// ---- 20_Module/Mqtt/Config/ST_ScheduleWeekly_V1.TcDUT
{attribute 'pack_mode' := '1'}
TYPE ST_ScheduleWeekly_V1 :
STRUCT
 Name : STRING(20);
 Priority : UDINT;
 StartDate : UDINT;
 EndDate : UDINT;
 Works : ARRAY[0..69] OF ST_ScheduleWork_V1;
END_STRUCT
END_TYPE

// ---- 20_Module/Mqtt/ST_IfUpsConfigRx.TcDUT
// MQTT로 받은 UPS 설정을 프로그램에 넘기는 묶음.
// 현재 수신만 하고 장비에는 적용하지 않는다.
{attribute 'pack_mode' := '1'}
TYPE ST_IfUpsConfigRx :
STRUCT
 nRxCount : UDINT; // 수신 누계
 astConfig : ARRAY[0..GVL_PARAM.UPS_COUNT-1] OF ST_UpsConfig_Rx; // UPS별 설정
END_STRUCT
END_TYPE

// ---- 20_Module/Ups/E_UpsChargeAction.TcDUT
// 충방전 시퀀스가 요청하는 동작. ST_UpsChargeRequest.eAction에 담긴다.
{attribute 'qualified_only'}
{attribute 'strict'}
TYPE E_UpsChargeAction : (
 NoRequest := 0, // 요청 없음
 BbcOn := 1, // BBC 기동
 BbcReady := 2, // BBC 대기 (현재 맵에 명령 없음, 확인 필요)
 BmsPreparePeriodic := 3, // BMS 주기적 방전 준비
 BmsPreparePulse := 4, // BMS 펄스 방전 준비
 PeriodicStart := 5, // UPS 주기적 방전 시작
 PulseStart := 6, // UPS 펄스 방전 시작
 DischargeCancel := 7, // UPS 방전 취소
 BmsDischargeCancel := 8, // BMS 방전 취소
 FloatCharge := 9, // 부동충전 복귀
 ChargeVoltage := 10 // 충전 전압 적용 (온도보상, fValue 사용)
) INT;
END_TYPE

// ---- 20_Module/Ups/E_UpsChargeMode.TcDUT
// 충방전 시퀀스의 운전 종류. 주 운전이라 한 번에 하나만 실행한다.
{attribute 'qualified_only'}
{attribute 'strict'}
TYPE E_UpsChargeMode : (
 Off := 0, // 운전 없음
 Trickle := 1, // 간헐충전
 Periodic := 2, // 주기적 방전
 Pulse := 3 // 펄스 방전
) INT;
END_TYPE

// ---- 20_Module/Ups/E_UpsChargeStep.TcDUT
// FB_UpsChargeSequence의 진행 단계.
{attribute 'qualified_only'}
{attribute 'strict'}
TYPE E_UpsChargeStep : (
 Idle := 0, // 대기
 WaitNormal := 10, // 시작 조건 확인
 WaitSchedule := 20, // 주기적 방전 일정 대기
 BbcStart := 30, // BBC 기동 요청
 WaitEnd := 40, // 종료 기준 도달 대기
 ExtraCharge := 50, // 추가 충전(간헐) / 초기 충전 대기(주기적)
 BbcReady := 60, // BBC 대기 요청
 WaitReady := 70, // BAT Mode 2 확인
 Rest := 80, // 휴지, 재충전 조건 대기
 PrepareBms := 90, // BMS 방전 준비 요청
 StartDischarge := 100, // UPS 방전 시작 요청
 WaitRunning := 110, // 방전 모드 진입 확인
 Running := 120, // 방전 실행 중
 CancelUps := 130, // UPS 방전 취소 요청
 CancelBms := 140, // BMS 방전 취소 요청
 BbcResume := 150, // 휴지 해제, BBC 재기동
 FloatRequest := 160, // 부동충전 요청
 WaitFloat := 170, // BAT Mode 0 확인
 Complete := 180, // 완료
 Fault := 900 // 고장 정지
) INT;
END_TYPE

// ---- 20_Module/Ups/ST_UpsChargeFeedback.TcDUT
// ST_UpsChargeRequest에 대한 처리 결과.
// nSeq가 요청 번호와 같고 bConfirmed가 TRUE여야 완료로 본다.
TYPE ST_UpsChargeFeedback :
STRUCT
 bValid : BOOL; // 확인 응답
 nSeq : UDINT; // 확인한 요청 번호
 bConfirmed : BOOL; // 동작 확인 완료
END_STRUCT
END_TYPE

// ---- 20_Module/Ups/ST_UpsChargeRequest.TcDUT
// 충방전 시퀀스가 장비 쪽에 보내는 요청 1건.
// nSeq로 요청을 구분하고, 처리 결과는 ST_UpsChargeFeedback으로 돌려받는다.
TYPE ST_UpsChargeRequest :
STRUCT
 bValid : BOOL; // 처리할 요청
 nSeq : UDINT; // 요청 번호
 eAction : E_UpsChargeAction; // 요청 동작
 fValue : REAL; // 전압 목표 (V)
END_STRUCT
END_TYPE

// ---- 20_Module/Ups/ST_UpsChargeSet.TcDUT
// 간헐충전·주기적 방전·펄스 방전·온도보상 설정값 묶음.
// 기본값은 예시이며 LiB 운전값은 미확정.
TYPE ST_UpsChargeSet :
STRUCT
 nTrickleCriterion : UINT; // 1: 전압, 2: SOC
 fStartVoltageV : REAL; // 재충전 시작 전압 (V)
 fEndVoltageV : REAL; // 추가충전 시작 전압 (V)
 fStartSocPct : REAL; // 재충전 시작 SOC (%)
 fEndSocPct : REAL; // 추가충전 시작 SOC (%)
 tExtraCharge : TIME := T#120M; // 추가 충전 시간
 tRestart : TIME := T#30D; // 대기 후 재충전 기간
 fFloatVoltageV : REAL; // 기준 부동충전 전압 (V)
 tInitialCharge : TIME := T#120M; // 주기적 방전 전 충전 시간
 fPeriodicCurrentA : REAL; // 주기적 방전 전류 (A)
 tPeriodicDischarge : TIME := T#10M; // 주기적 방전 시간
 wMonthMask : WORD; // 1~12월 선택 비트 0~11
 nWeek : UINT; // 월내 1~4주차 (1~7일이 1주차)
 nWeekDay : UINT; // 0: 일요일 ~ 6: 토요일
 nHour : UINT; // 실행 시간 (0~23)
 fPulseChargeA : REAL; // 펄스 충전 전류 (A)
 fPulseDischargeA : REAL; // 펄스 방전 전류 (A)
 tPulseCharge : TIME := T#5S; // 펄스 충전 시간
 tPulseDischarge : TIME := T#5S; // 펄스 방전 시간
 nPulseCycles : UINT; // DSP 실행 횟수
 tRunTimeout : TIME := T#1H; // 방전 완료 감시 시간
 tRequestTimeout : TIME := T#10S; // 요청 확인 대기 시간
 tModeTimeout : TIME := T#30S; // 운전 모드 확인 대기 시간
 fBaseCellVoltageV : REAL; // 25℃ 기준 셀 전압 (V)
 nSeriesCells : UINT; // 직렬 셀 수
 fSlopeMvPerC : REAL; // 셀당 온도 기울기 (mV/℃)
 fMinChargeVoltageV : REAL; // 적용 가능한 최저 전압 (V)
 fMaxChargeVoltageV : REAL; // 적용 가능한 최고 전압 (V)
 fMinTemperatureC : REAL; // 보상 가능한 최저 온도 (℃)
 fMaxTemperatureC : REAL; // 보상 가능한 최고 온도 (℃)
 tTempUpdate : TIME := T#1M; // 온도보상 갱신 주기
END_STRUCT
END_TYPE

// ---- 20_Module/Ups/ST_UpsDesiredSet.TcDUT
(* UPS 1대에 맞춰 둘 설정 보관값 (장치: UPS). 2026-11-05.
   기반 없음(신규). GVL_PERSIST.g_astUpsDesired에 두어 PMS 재시작 후에도 남는다.
   명세: C:\gil\UPS\명세서\UPS_명세서.md CF-UPS-02·03
   칸 0~6 = UPS Holding H50~H56 (FB_UpsConfigApply의 쓰기 대상과 같은 순서)
   bTempCompOn·bTrickleOn = 시작·정지 명령으로 정한 켜짐 상태 (FB_UpsCommand가 씀, 2026-11-05 추가) *)
TYPE ST_UpsDesiredSet :
STRUCT
	bValid		: BOOL;							// 한 번이라도 EMS 설정을 받아 보관함
	abUse		: ARRAY[0..6] OF BOOL;			// 이 칸을 맞출지 (EMS is_available)
	awValue		: ARRAY[0..6] OF WORD;			// 맞출 원시값 (UPS 레지스터 값 그대로)
	nRxCount	: UDINT;						// 보관한 설정의 수신 누계 (참고용)
	bTempCompOn	: BOOL;							// 온도보상충전을 켜 둬야 함 (명령 4 → TRUE, 8 → FALSE)
	bTrickleOn	: BOOL;							// 간헐충전을 켜 둬야 함 (명령 1 → TRUE, 7 → FALSE). UPS 상태로 확인할 칸이 없어 복구는 하지 않음
END_STRUCT
END_TYPE

// ---- 20_Module/Ups/ST_IfUpsCmd.TcDUT
(* EMS UPS 명령 1건 (MqttTask → PlcTask 칸, GVL_IF.g_astUpsCmd). 2026-11-05. 명세: WR-UPS-01 *)
TYPE ST_IfUpsCmd :
STRUCT
	nSeq	: UDINT;	// 새 명령마다 1씩 오름. 받는 쪽은 번호 변화로 새 명령을 안다
	nType	: UDINT;	// 명령 번호 1~26 (EMS CommandType 그대로. 인터페이스 100.Command, 명세 WR-UPS-01)
END_STRUCT
END_TYPE

// ---- 20_Module/Driver/LS/ST_LsImd1000State.TcDUT
(* LS IMD1000 읽은 값 (FB_LsImd1000.q_stState → FB_RptLsImd1000). 2026-11-09.
   맵: 인터페이스\(MM-20210721) IMD1000 Modbus-Setting_v1_0_0.pdf 3.6.2·3.6.3. 주소는 프로토콜 주소(0 기준, 맵 Addr 열) *)
TYPE ST_LsImd1000State :
STRUCT
	bValid		: BOOL;		// 통신 정상이고 측정 영역을 한 번 이상 읽음
	fInsulation	: REAL;		// 절연저항 kΩ (IR 224~225 FLOAT32, 앞 = 상위 워드)
	wDiState	: WORD;		// IR 206 기기 DI 입력 상태 (b0 버튼 Self Test, b1 DI Self Test, b2 DI Stand-By)
	wSelfDiag	: WORD;		// IR 209 자가진단-기기 Error 상태#2 (b0 메모리, b1 RTC, b2 교정)
	wAlarm		: WORD;		// IR 210 절연저항 측정 alarm 상태 (b0 Ins. Alarm, b1~b3 Pre Alarm#1~#3 동작)
	wConnect	: WORD;		// IR 211 기기 & 계통 연결 상태 (b0 PE 연결, b1 Device, b2 System 연결, b8 측정 전압 이상)
	wSelfTest	: WORD;		// IR 215 Self Test 전체 진행 상태 (0 없음, 1 진행, 2 완료, 5 정지)
	bSetValid	: BOOL;		// 설정 영역을 한 번 이상 읽음
	nInsPickup	: UDINT;	// HR 40~41 Ins. Alarm Pick-up kΩ (UINT32, 앞 = 상위 워드)
	nPre1Pickup	: UDINT;	// HR 46~47 Pre Alarm#1 Pick-up kΩ
END_STRUCT
END_TYPE

// ---- 20_Module/Common/ST_TempHumState.TcDUT
(* 온습도계 읽은 값 (드라이버 q_stState → FB_RptTempHum → 토픽 temperature_sensor). 2026-11-09.
   ITGuard IE-SX·RADIONODE RN172 같이 씀 *)
TYPE ST_TempHumState :
STRUCT
	bValid		: BOOL;		// 통신 정상이고 센서 값이 유효
	fTemp		: REAL;		// 온도 ℃
	fHum		: REAL;		// 습도 %
END_STRUCT
END_TYPE

// ---- 20_Module/Mqtt/Publish/ST_ImdPublish_V1.TcDUT
(* EMS로 보내는 IMD 레코드 1개 (토픽 imd). 인터페이스\22. IMD.xlsx V1 그대로, 32 B. 바이너리 구조라 필드 순서를 바꾸면 안 된다. 2026-11-09 *)
{attribute 'pack_mode' := '1'}
TYPE ST_ImdPublish_V1 :
STRUCT
	DeviceIndex							: UDINT;	// 장치 번호 (1부터)
	Status								: UDINT;	// b0 통신에러, b1 Pre-Warning, b2 Warning, b3 Fault, b4 Alarm, b5 Internal test, b6 External test
	InsulationResistance				: REAL;		// 절연저항 kΩ
	DeviceErrorLocation					: REAL;		// 에러난 장치의 Device Number (Bender 항목, IMD1000은 0)
	InsulationResistanceFaultLocation	: REAL;		// 0~25 (+)극, 75~100 (-)극 (Bender 항목, IMD1000은 0)
	PreAlarmSettingValue				: UDINT;	// 사전경보 설정값 kΩ
	MainAlarmSettingValue				: UDINT;	// 주경보 설정값 kΩ
	Fault1								: UDINT;	// b0 SystemConnection Error, b1 ConnectionToEarth Error
END_STRUCT
END_TYPE

// ---- 20_Module/Mqtt/Publish/ST_ImdPublishData.TcDUT
(* EMS로 보내는 IMD MQTT 패킷 전체 (토픽 imd). 바이너리 구조라 필드 순서를 바꾸면 안 된다. 2026-11-09 *)
{attribute 'pack_mode' := '1'}
TYPE ST_ImdPublishData :
STRUCT
	Header		: ST_MqttHeader;									// MQTT 공통 헤더
	Devices		: ARRAY[0..GVL_PARAM.IMD_COUNT-1] OF ST_ImdPublish_V1;	// IMD별 데이터
END_STRUCT
END_TYPE

// ---- 20_Module/Mqtt/Publish/ST_FirePublish_V1.TcDUT
(* EMS로 보내는 화재감지기 레코드 1개 (토픽 fire_detector, 이름 잠정). 인터페이스 20. OffGas.xlsx V1과 같은 모양, 8 B. 2026-11-10 사용자 결정
   바이너리 구조라 필드 순서를 바꾸면 안 된다 *)
{attribute 'pack_mode' := '1'}
TYPE ST_FirePublish_V1 :
STRUCT
	DeviceIndex	: UDINT;	// 장치 번호 (1부터: 1 = TS-60, 2 = ASD-57. UPSstd 번호 규칙)
	Status		: UDINT;	// b0 통신 이상, b1 알람 (연기 등 감지), b2 고장 (감지기 자체 이상, 알 수 있을 때만)
END_STRUCT
END_TYPE

// ---- 20_Module/Mqtt/Publish/ST_FirePublishData.TcDUT
(* EMS로 보내는 화재감지기 MQTT 패킷 전체 (토픽 fire_detector, 이름 잠정). 바이너리 구조라 필드 순서를 바꾸면 안 된다. 2026-11-10 *)
{attribute 'pack_mode' := '1'}
TYPE ST_FirePublishData :
STRUCT
	Header		: ST_MqttHeader;										// MQTT 공통 헤더
	Devices		: ARRAY[0..GVL_PARAM.FIRE_COUNT-1] OF ST_FirePublish_V1;	// 감지기별 데이터
END_STRUCT
END_TYPE

// ---- 20_Module/Driver/Esolution/ST_BatRackCmd.TcDUT
(* EMS 랙 컨택터 명령 하나 (command/bat CommandType 11 닫기, 12 열기, Value = 랙 번호). 2026-11-10.
   쓰는 곳: FB_EmsCommand, 읽는 곳: MAIN → FB_BmsRackCommand. 명세 WR-BAT-01 *)
TYPE ST_BatRackCmd :
STRUCT
	nSeq		: UDINT;	// 명령 번호. 바뀌면 새 명령 (0 = 한 번도 못 받음)
	nRack		: UINT;		// 랙 번호 1~ (BMS 안 번호). 범위 밖이면 거절
	bClose		: BOOL;		// TRUE = 랙 닫기(11), FALSE = 랙 열기(12)
END_STRUCT
END_TYPE

// ---- 20_Module/Driver/Esolution/ST_BatCtlCmd.TcDUT
(* EMS 컨택터 하나씩 명령 (command/bat CommandType 5~10). 2026-11-13.
   5 시스템(랙 전체 40013) 연결, 6 차단, 7 충전 컨택터(40014) 닫기, 8 열기, 9 방전 컨택터(40015) 닫기, 10 열기
   쓰는 곳: FB_EmsCommand, 읽는 곳: MAIN → FB_BmsContactorCommand. 인터페이스 100.Command BAT *)
TYPE ST_BatCtlCmd :
STRUCT
	nSeq		: UDINT;	// 명령 번호. 바뀌면 새 명령 (0 = 한 번도 못 받음)
	nType		: UINT;		// CommandType 5~10 (그 밖은 거절)
END_STRUCT
END_TYPE

// ---- 10_Core/00_Type/GVL_REASON.TcGVL
VAR_GLOBAL CONSTANT
	(* 코어가 낸 제한의 이유 코드 (모듈 ID = 0일 때)
	   - 모듈 ID ≠ 0이면 이유 코드는 그 모듈이 정한 것. 지령원이 낸 제한은 이유 0 *)
	RSN_RATING		: UINT := 1;		// 가용 유닛 P 정격 합
	RSN_BAT			: UINT := 2;		// 배터리 충·방전 한도 합
	RSN_RATING_Q	: UINT := 3;	// 가용 유닛 Q 정격 합
	RSN_DERATE	: UINT := 4;	// 보호 Derate (유닛 정격 × Derate)
END_VAR

// ---- 10_Core/00_Type/GVL_CORE.TcGVL
VAR_GLOBAL CONSTANT
	(* 코어 내부 상수 (현장에서 바꾸지 않음. 현장 대수·크기는 GVL_PARAM) *)
	NO_LIMIT		: REAL := 1.0E9;	// 정격·배터리가 없어 한도를 걸 수 없는 유닛·버스의 대용 한도 (kW·kvar). 열린 범위·무한대 판정(F_RangeOpen·F_CmdOk)의 1E30과는 뜻이 다름
END_VAR

// ---- 90_Project/GVL_TEST.TcGVL
VAR_GLOBAL
	g_astVirtual	: ARRAY[1..GVL_PARAM.GROUP_COUNT] OF ST_VirtualSet;	// 가상신호. 저장 안 함 (재기동 시 꺼짐)
	g_bTestReset	: BOOL;		// 시험: 모든 PCS·BMS 고장 리셋 명령 + 유지 DO 풀기 (TEST_MODE에서만)
END_VAR

// ---- 90_Project/GVL_MQTT.TcGVL
VAR_GLOBAL CONSTANT
	(* ================================================================
	   MQTT 보고·명령 (PMS ↔ EMS 토탈 인터페이스)
	   - 장치 수는 GVL_PARAM (PCS_COUNT, BMS_COUNT, RACK_COUNT, PV_COUNT, ESS_COUNT, TEMP_COUNT, AIR_CONDITIONER_COUNT)
	   - 토픽: 발행 dgspms/{SOLUTION_NAME}/{사이트}/{장치} , config echo dgspms/.../config/{장치}
	           구독 dgsems/{SOLUTION_NAME}/{사이트}/{command|config}/{장치}
	           로거 dgspms/{SOLUTION_NAME}/{사이트}/pms_log (이벤트 로그, 발생할 때 1건씩. 20_Module/Mqtt/Logger)
	   - 접속 설정(사이트 번호·브로커 주소·포트·계정)은 GVL_SITE.MQTT_SET
	   ================================================================ *)
	DEVICE_TOPIC_COUNT	: UINT := 12;		// 발행 장치 토픽 수: pms pcs bat rack pv ess temp airconditioner ups module imd fire_detector
	CONFIG_TOPIC_COUNT	: UINT := 4;		// config 토픽 수: pcs bat protection ups (구독, 받은 값 echo 발행)
	COMMAND_TOPIC_COUNT	: UINT := 3;		// command 토픽 수: pcs bat ups (구독). ups는 2026-11-05 추가 (명세 WR-UPS-01)
	UPS_REPORT_ENABLED : BOOL := TRUE; // FB_RptSebangUps 매핑 연결됨
	IMD_REPORT_ENABLED : BOOL := TRUE; // FB_RptLsImd1000 매핑 연결됨 (인터페이스 22. IMD)
	FIRE_REPORT_ENABLED : BOOL := TRUE; // 화재감지기 보고 (fire_detector, 토픽 이름 잠정. 인터페이스 20. OffGas 양식)
	MODULE_REPORT_ENABLED : BOOL := TRUE; // 시험: BMS1 시뮬레이터. 모듈 레코드에 유효 표시가 없어 무효 데이터는 0, Rack Status b0로 구분
	SOLUTION_NAME		: STRING(15) := 'ups';		// 토픽 두 번째 칸 (모든 토픽에 들어감)

	HEADER_VERSION		: UDINT := 1;
	DEVICE_VERSION		: UDINT := 1;
	COMMAND_VERSION		: UDINT := 2;

	(* 로거 (이벤트 로그 → pms_log 토픽). 메시지 1건 = 이벤트 1건 (ST_LoggerPublish_V1) *)
	LOGGER_TOPIC		: STRING(15) := 'pms_log';
	LOGGER_VERSION		: UDINT := 1;		// 로거 패킷 헤더 DeviceVersion
	LOGGER_QUEUE		: UINT := 64;		// 이벤트 큐 칸 수 (브로커가 끊기거나 접속 전인 동안 이만큼 보관. 한 스캔에 생길 수 있는 로그 수보다 커야 함: PRG_TestLogger.bSendAll은 스캔마다 32건)
	LOGGER_TEXT_MAX		: INT := 100;		// Contents 글자 수. ST_LoggerPublish_V1.Contents·ST_LoggerSlot.wsText의 WSTRING(100)과 같게 (로그 문구 규칙 95자 + 해소 표시 5자)
	LOGGER_LANG_ID		: DINT := 1033;		// 이벤트 문구를 요청할 언어. 문구는 기본 언어 하나뿐이라 이 값으로 그 문구가 옴 (시험 때 확인)
END_VAR

VAR_GLOBAL
	(* ---------- 발행 패킷 (헤더 + 장치 배열). 장치 배열은 0부터 = 레코드 DeviceIndex(RACK DeviceID) = DB 장치키 ---------- *)
	g_stPmsPublish			: ST_PmsPublishData;
	g_stPcsPublish			: ST_PcsPublishData;
	g_stBatPublish			: ST_BatPublishData;
	g_stRackPublish			: ST_RackPublishData;
	g_stUpsPublish : ST_UpsPublishData;
	g_stModulePublish : ST_ModulePublishData;
	g_stImdPublish			: ST_ImdPublishData;		// IMD (절연감시)
	g_stFirePublish			: ST_FirePublishData;		// 화재감지기 (연기)
	g_stPvPublish			: ST_PvPublishData;
	g_stEssPublish			: ST_EssPublishData;
	g_stTempPublish			: ST_TempPublishData;
	g_stAirConditionerPublish	: ST_AirConditionerPublishData;	// 공조기

	(* ---------- 구독 수신 (받은 레코드를 장치 번호 칸에 넣음. 받은 DeviceIndex 0 → 칸 0, F_MqttDistribute.DEVICE_ID_BASE) ---------- *)
	g_astPcsCommand			: ARRAY[0..GVL_PARAM.PCS_COUNT-1] OF ST_MqttCommand_Rx;	// command/pcs. FB_EmsCommand가 처리 후 CommandType을 0으로 지움
	g_astBatCommand			: ARRAY[0..GVL_PARAM.BMS_COUNT-1] OF ST_MqttCommand_Rx;	// command/bat
	g_astUpsCommand			: ARRAY[0..GVL_PARAM.UPS_COUNT-1] OF ST_MqttCommand_Rx;	// command/ups (DeviceIndex 1부터). PRG_Mqtt가 GVL_IF.g_astUpsCmd로 넘기고 CommandType을 0으로 지움
	g_astPcsConfig			: ARRAY[0..GVL_PARAM.PCS_COUNT-1] OF ST_PcsConfig_Rx;		// config/pcs
	g_astBatConfig			: ARRAY[0..GVL_PARAM.BMS_COUNT-1] OF ST_BatConfig_Rx;		// config/bat
	g_astUpsConfig : ARRAY[0..GVL_PARAM.UPS_COUNT-1] OF ST_UpsConfig_Rx; // received values only, not approved settings
	g_stUpsConfigWireIn : ST_UpsConfigWirePacket;
	g_stUpsConfigEcho : ST_UpsConfigWirePacket; // receipt echo, NEVER means device applied
	g_stProtectionConfig	: ST_ProtectionConfig_Rx;										// config/protection

	(* config 수신 버퍼 (헤더 + 레코드). 헤더의 Location·UserName을 echo에 그대로 씀 *)
	g_stPcsConfigWireIn			: ST_PcsConfigWirePacket;
	g_stBatConfigWireIn			: ST_BatConfigWirePacket;
	g_stProtectionConfigWireIn	: ST_ProtectionConfigWirePacket;

	(* config echo 발행 패킷 *)
	g_stPcsConfigEcho		: ST_PcsConfigWirePacket;
	g_stBatConfigEcho		: ST_BatConfigWirePacket;
	g_stProtectionConfigEcho	: ST_ProtectionConfigWirePacket;	// [결함 12 수정 2026-11-04: 추가. 원래 g_stProtectionConfigWireIn을 그대로 발행했는데 아무도 안 채워 0으로 나감]

	(* 수신 기록 (3개 브로커 합산) *)
	g_asCmdRxTime			: ARRAY[1..GVL_MQTT.COMMAND_TOPIC_COUNT] OF STRING(23);	// 토픽별 마지막 command 헤더 TimeStamp
	g_asCfgRxTime			: ARRAY[1..GVL_MQTT.CONFIG_TOPIC_COUNT] OF STRING(23);
	g_anCmdRxCount			: ARRAY[1..GVL_MQTT.COMMAND_TOPIC_COUNT] OF UDINT;		// 토픽별 새 command 수신 횟수
	g_anCfgRxCount			: ARRAY[1..GVL_MQTT.CONFIG_TOPIC_COUNT] OF UDINT;
	g_anCfgRxRecords		: ARRAY[1..GVL_MQTT.CONFIG_TOPIC_COUNT] OF UDINT;	// 토픽별 마지막 새 메시지에서 실제로 받은 레코드 수 (PRG_Mqtt가 빈 칸과 '모두 is_available 0' 레코드를 구분) [21번 수정 2026-11-09: 추가]
	(* 실제 반영된 config (MAIN → GVL_IF → PRG_Mqtt). FB_MqttMain이 echo로 발행. 아직 못 받았으면(g_bConfigApplied FALSE) 받은 값을 echo [9-21 수정 2026-11-04: 추가] *)
	g_astPcsConfigApplied	: ARRAY[0..GVL_PARAM.PCS_COUNT-1] OF ST_PcsConfig_Rx;
	g_astBatConfigApplied	: ARRAY[0..GVL_PARAM.BMS_COUNT-1] OF ST_BatConfig_Rx;
	g_bConfigApplied		: BOOL;
END_VAR

// ---- 20_Module/ControlMode/GVL_CM_RSN.TcGVL
{attribute 'qualified_only'}
VAR_GLOBAL CONSTANT
	(* 요금제 기반 제어 모드(FB_CmTariffBase 파생)의 상태·이유 코드. 문구는 FB_CmTariffBase.M_ReasonText
	   q_nState: 0 = 정상(값 그대로), 아래 = 지금 출력이 왜 이런지. M_CheckEnter·bExitReq의 이유 코드도 같은 표 *)
	NO_TIME		: UINT := 1;	// 시각 무효 → 0 (진입 거부)
	NO_UNIT		: UINT := 2;	// 가용 유닛 없음 (진입 거부)
	HOLIDAY		: UINT := 3;	// 휴일 → 0
	NO_SLOT		: UINT := 4;	// 맞는 시간표 칸 없음 → 0
	DIS_TIME	: UINT := 5;	// 방전 허용 시간 아님 → 0
	REV_LIMIT	: UINT := 6;	// 역송 방지로 방전을 줄임
	NO_PCC		: UINT := 7;	// 접속점 계측 무효 → 방전 0
	NO_CAP		: UINT := 8;	// 배터리 용량·SOC 무효 → 0
	PEAK		: UINT := 11;	// 피크 제어 방전
	BELOW_PEAK	: UINT := 12;	// 피크 제어 필요 없음 → 0
	AUTO_CHG	: UINT := 13;	// 자동 충전 시간
	REMAIN_DIS	: UINT := 14;	// 잔량 방전 시간
	SCHED_PEAK	: UINT := 15;	// 스케줄 방전과 피크 제어 중 큰 값
	NEW_INTERVAL: UINT := 16;	// 새 15분 구간 첫 스캔 → 0
END_VAR

// ---- 90_Project/GVL_PARAM.TcGVL
VAR_GLOBAL CONSTANT
	(* ================================================================
	   대수·크기 (라이브러리로 나누면 라이브러리 파라미터 리스트가 됨)
	   - 코어와 모듈은 GVL_SITE·GVL_PERSIST를 보지 않고 이 값만 쓴다.
	   - 등록 칸 수는 최소 1. 비워 둔 칸은 "등록 안 함"으로 본다.
	   - 값을 바꾸면 배열 크기가 바뀌므로 재빌드·액티베이트.
	   ================================================================ *)

	(* ---------- 장비 ---------- *)
	INSTALLED_PCS_COUNT : UINT := 0; // no separate PCS in this UPS site; allocation slots remain below
	PCS_COUNT		: UINT := 2;		// PCS 대수
	MAX_SUB			: UINT := 1;		// PCS 1대 안에서 따로 제어하는 유닛 최대 수
	UNIT_COUNT		: UINT := 2;		// 제어 유닛 수 (구성은 GVL_SITE.UNIT_CFG)
	BMS_COUNT		: UINT := 1;		// BMS 장비 수 (현장 5: BAT 1대) (소속 배터리 그룹은 GVL_SITE.BMS_CFG)
	BAT_COUNT		: UINT := 1;		// 배터리 그룹(DC 버스) 수 (현장 5: 1). 유닛 n : BMS m을 한 그룹으로 묶음
	METER_COUNT		: UINT := 1;		// 계측기 수
	AUX_COUNT		: UINT := 7;		// 보조 장비 칸 수 (GVL_SITE.g_aipAux: 1 온습도(오토닉스), 2 IMD(LS IMD1000), 3 원격 I/O, 4 온습도(ITGuard), 5 지락검출계전기, 6 벡호프 단자 I/O(TS-60), 7 ASD-57 감지기)
	AUX_DI_MAX		: UINT := 16;		// FB_AuxIo 하나의 점 수: 디지털 입력
	AUX_DO_MAX		: UINT := 16;		// 디지털 출력
	AUX_AI_MAX		: UINT := 8;		// 아날로그 입력
	AUX_AO_MAX		: UINT := 4;		// 아날로그 출력

	(* ---------- 보고(MQTT)만 하는 장치 (제어하지 않음). PCS·BAT 보고 수는 PCS_COUNT·BMS_COUNT ---------- *)
	UPS_ALGORITHM_ENABLED : BOOL := FALSE; // 충방전 로직 기본 차단
	UPS_CONTROL_ENABLED : BOOL := FALSE; // code-only gate for ALL new UPS/BMS hardware writes
	UPS_CFG_MAX_CURRENT_A : REAL := 100.0; // EMS 방전·펄스 전류 상한 (A). 시험값, 운전값 확정 시 변경
	UPS_CFG_MAX_MINUTES : UDINT := 60; // EMS 주기적 방전 시간 상한 (분)
	UPS_CFG_MAX_SECONDS : UDINT := 60; // EMS 펄스 시간 상한 (초)
	UPS_CFG_MAX_CYCLES : UDINT := 1000; // EMS 펄스 횟수 상한
	UPS_COUNT		: UINT := 1;		// UPS 대수 (현장 5: 1대). PCS와 별개이며 실제 드라이버는 미연결
	RACKS_PER_BMS	: UINT := 8;		// 배터리 시스템 한 대당 랙 수 (현장 5: 8, 드라이버 최대 10)
	MODULES_PER_RACK : UINT := 9;		// 랙 한 개당 배터리 모듈 수 (현장 5: 9, 맵 최대 17)
	CELLS_PER_MODULE : UINT := 14;		// 모듈 한 개당 셀 수 (현장 5: 14). BMS 맵은 모듈당 셀 20칸, MQTT module 레코드도 CellVoltage1~20 그대로 (15~20은 0)
	RACK_COUNT		: UINT := BMS_COUNT * RACKS_PER_BMS;	// MQTT rack 레코드 총 8개
	BAT_MODULE_COUNT : UINT := RACK_COUNT * MODULES_PER_RACK;	// 배터리 모듈 총 72개 (PLC 기능 모듈 수 MODULE_MAX와 별개)
	PV_COUNT		: UINT := 1;		// PV 수 (MQTT pv_meter 토픽)
	ESS_COUNT		: UINT := 1;		// ESS 수 (MQTT ess_meter 토픽)
	TEMP_COUNT		: UINT := 1;		// 온도 장치 수 (MQTT temperature_sensor 토픽)
	IMD_COUNT		: UINT := 1;		// IMD(절연감시) 수 (MQTT imd 토픽). MAIN.A_Report가 칸마다 GVL_SITE.g_fbImdN을 연결
	FIRE_COUNT		: UINT := 2;		// 화재감지기 수 (MQTT fire_detector 토픽, OffGas 양식). 1 = TS-60 연기 접점, 2 = ASD-57
	AIR_CONDITIONER_COUNT	: UINT := 1;	// 공조기 수 (MQTT airconditioner 토픽)

	(* ---------- 계측점 ---------- *)
	POINT_COUNT		: UINT := 1;		// 계측점 수 (구성은 GVL_SITE.POINT_CFG)
	POINT_TERM_MAX	: UINT := 3;		// 계측점 하나에 묶는 계측기 최대 수

	(* ---------- 제어 그룹 ---------- *)
	GROUP_COUNT		: UINT := 1;		// 제어 그룹 수 (접속점 1개 + 소속 유닛)

	(* ---------- 모듈 등록 칸 수 ---------- *)
	SOURCE_COUNT	: UINT := 3;		// 지령원. 1 = 시험, 2 = 제어 모드 관리자 (접속점 그룹 1), 3 = EMS [16번 수정 2026-11-09: 원래 4 (2 = 관리자 PCS1, 3 = 관리자 PCS2, 4 = EMS)]
	LIMIT_COUNT		: UINT := 1;		// 출력 제한
	PERMIT_COUNT	: UINT := 1;		// 기동 조건
	COMP_COUNT		: UINT := 1;		// 보정
	RULE_COUNT		: UINT := 7;		// 보호 규칙 (1~5 = 표준 보호 5종, 현장 보호는 6부터. 6 = 연기 TS-60, 7 = 연기 ASD-57)
	OUTPUT_COUNT	: UINT := 1;	// 출력 규칙 (보조 장비 DO: 팬·경광등·트립 등)
	UNIT_RULE_COUNT	: UINT := 1;	// 유닛 제한 (사용자 한도 등)
	BAT_RULE_COUNT	: UINT := 1;	// 버스 제한 (SOC 감발 등)
	CTRL_MODE_COUNT	: UINT := 5;	// 제어 모드 (FB_CtrlModeMgr 하나에 등록하는 모드 수. 한 번에 하나만 켬. 틀은 10_Core, 모드는 20_Module\ControlMode). 1 = 정출력, 2 = 스케줄, 3 = 피크컷, 4 = 통합, 5 = 스탠다드 스케줄(EMS 지령). 관리자는 PCS마다 하나 (GVL_SITE)
	SCHED_SLOT_COUNT	: UINT := 10;	// 스케줄 모드 시간표 칸 수 (계절·요일마다)
	MODULE_SET_BYTES	: UDINT := 8192;	// 현장 모듈 설정 묶음(GVL_PERSIST.g_stModuleSet) 최대 크기. 넘으면 바뀌어도 바로 저장 안 됨 (fbPersistSave.q_bModuleSetTooBig)

	(* ---------- 계산값 (고치지 않음) ---------- *)
	MODULE_MAX		: UINT := PCS_COUNT + BMS_COUNT + METER_COUNT + AUX_COUNT + SOURCE_COUNT + LIMIT_COUNT + PERMIT_COUNT + COMP_COUNT + 2 * RULE_COUNT + OUTPUT_COUNT + UNIT_RULE_COUNT + BAT_RULE_COUNT + 2 * GROUP_COUNT + 2;	// 뒤 = 그룹별 고르기·분배 정책, Auto·Manual Gate
	PROT_TARGET_MAX	: UINT := UNIT_COUNT + BMS_COUNT + BAT_COUNT + GROUP_COUNT;	// 보호 규칙 하나가 보는 대상 번호 상한 (범위마다 대상 수가 달라 넉넉하게 합)
	TRACE_STEP_MAX	: UINT := 8 + 2 * LIMIT_COUNT;		// 출력 추적표 줄 수: 요청·램프·보정·정격·배터리·분배 후·쓴 값 + 지령원 제한 + 제한 모듈마다 (접속점·설비)
END_VAR

// ---- 90_Project/GVL_PERSIST.TcGVL
VAR_GLOBAL PERSISTENT
	(* ================================================================
	   운영 설정 (HMI에서 바꿈, 재기동 후에도 유지)
	   - 칸 순서는 GVL_SITE 등록 배열과 같다
	   - 설정을 추가하면 MAIN.fbPersistSave에도 연결한다 (바뀌면 바로 저장)
	   ================================================================ *)
	g_aeOpMode		: ARRAY[1..GVL_PARAM.UNIT_COUNT] OF E_OpMode;	// 유닛별 운전 모드 요청 (HMI가 쓰고, 보호가 ToManual이면 FB_ModeSwitch가 Manual로 바꿈). 실제 모드는 MAIN.fbModeSwitch.q_aeOpMode
	g_astGroupSet	: ARRAY[1..GVL_PARAM.GROUP_COUNT] OF ST_GroupSet;	// 제어 그룹별 선택 방식·램프·Q 필터
	g_astManualPolicy: ARRAY[1..GVL_PARAM.GROUP_COUNT] OF ST_ManualPolicy;	// 제어 그룹별 Manual 경로에 적용할 단계 (운전 정책·장비 보호 켜고 끄기)

	g_astSourceReg	: ARRAY[1..GVL_PARAM.SOURCE_COUNT] OF ST_SourceReg := [
						(bEnable := TRUE, nGrade := 1, stStateMode := (stPcs := (eRun := E_SourceMode.Both, eStandby := E_SourceMode.Both, eStop := E_SourceMode.Both, eEStop := E_SourceMode.Both), stBat := (eClose := E_SourceMode.Both, eOpen := E_SourceMode.Both)), ePowerMode := E_SourceMode.Both, nGroup := 0, tExpire := T#10S),	// 1 시험 지령원 (상태·출력 모두 Auto·Manual에서 받음)
						(bEnable := TRUE, nGrade := 2, stStateMode := (stPcs := (eRun := E_SourceMode.None, eStandby := E_SourceMode.None, eStop := E_SourceMode.None, eEStop := E_SourceMode.None), stBat := (eClose := E_SourceMode.None, eOpen := E_SourceMode.None)), ePowerMode := E_SourceMode.Auto, nGroup := 0, tExpire := T#10S),	// 2 제어 모드 관리자 접속점 그룹 1 (Auto 유닛 P·Q만, 상태 요청 안 받음) [16번 수정 2026-11-09: 원래 2 = 관리자 PCS1, 3 = 관리자 PCS2]
						(bEnable := TRUE, nGrade := 2, ePowerMode := E_SourceMode.Auto, nGroup := 0, tExpire := T#60S, bLostAlarm := FALSE,
							stStateMode := (stPcs := (eRun := E_SourceMode.Auto, eStandby := E_SourceMode.Auto, eStop := E_SourceMode.Both, eEStop := E_SourceMode.Both),
											stBat := (eClose := E_SourceMode.Auto, eOpen := E_SourceMode.Auto)))];	// 3 EMS [9번 수정 2026-11-09: bLostAlarm FALSE — '지령원 끊김' 대신 '브로커 끊김' 알람 (g_stBrokerWatch)] (상태 명령은 Auto에서 받고 정지·비상정지는 Manual에서도 받음. P 지령은 FB_SrcEms.i_bPEnable이 켜질 때만. EMS가 60 s 안에 다시 말하지 않으면 끊김)
	g_astLimitReg	: ARRAY[1..GVL_PARAM.LIMIT_COUNT] OF ST_ModuleReg;
	g_astPermitReg	: ARRAY[1..GVL_PARAM.PERMIT_COUNT] OF ST_ModuleReg;
	g_astCompReg	: ARRAY[1..GVL_PARAM.COMP_COUNT] OF ST_ModuleReg;
	g_astRuleCfg	: ARRAY[1..GVL_PARAM.RULE_COUNT] OF ST_RuleCfg := [	// 보호 규칙 (칸 = GVL_SITE.g_aipRule·g_aipResp). nTarget 0 = 범위 안 대상 전부. stProt 조치는 표준 대응(대응 칸에 g_fbProtRespStd)이 씀. 대응 칸이 비면 조치 없음 ([결함 8 수정 2026-11-03: 주석 고침. 원래 '표준 대응(대응 칸이 빈 칸)이 씀'])
						(stProt := (ePcsAction := E_PcsAction.Stop), eScope := E_ProtScope.Unit),		// 1 PCS 고장 → 그 유닛 정지
						(stProt := (ePcsAction := E_PcsAction.Standby), eScope := E_ProtScope.Unit),	// 2 PCS 통신 끊김 → 그 유닛 대기
						(stProt := (ePcsAction := E_PcsAction.Stop, eBatAction := E_BatAction.Stop), eScope := E_ProtScope.Bms),	// 3 BMS 고장 → 그 BMS 정지 + 같은 배터리 그룹 유닛 정지
						(stProt := (ePcsAction := E_PcsAction.Standby), eScope := E_ProtScope.Bms),		// 4 BMS 통신 끊김 → 같은 배터리 그룹 유닛 대기
						(stProt := (ePcsAction := E_PcsAction.Standby), eScope := E_ProtScope.Group),	// 5 접속점 계측 무효 → 그룹 대기
						(stProt := (ePcsAction := E_PcsAction.None), eScope := E_ProtScope.Site),		// 6 연기 감지 (TS-60) → 알람만
						(stProt := (ePcsAction := E_PcsAction.None), eScope := E_ProtScope.Site)];		// 7 연기 감지 (ASD-57) → 알람만
						(* BMS 하나가 빠져도 남은 BMS로 계속 돌리려면 3·4번 ePcsAction을 None으로 (3번은 eBatAction도 None: 배터리 조치는 PCS 정지·비상정지와만) *)
	g_astOutputCfg	: ARRAY[1..GVL_PARAM.OUTPUT_COUNT] OF ST_OutputCfg;	// 출력 규칙 (어느 장비·점, 임계값, 지연, 유지)
	g_astUnitRuleReg	: ARRAY[1..GVL_PARAM.UNIT_RULE_COUNT] OF ST_RuleTargetReg;	// 유닛 제한 모듈 등록 (대상 유닛, 적용 운전 모드)
	g_astBatRuleReg	: ARRAY[1..GVL_PARAM.BAT_RULE_COUNT] OF ST_RuleTargetReg;	// 버스 제한 모듈 등록 (대상 배터리 그룹, 적용 운전 모드). 1 = SOC 정책 (기본: 전체 버스, Auto·Manual)

	(* UPS 설정 보관값 (명세 CF-UPS-02). EMS에서 받은 설정. FB_UpsConfigApply가 쓰고, 바뀌면 fbPersistSave가 바로 저장 *)
	g_astUpsDesired	: ARRAY[1..GVL_PARAM.UPS_COUNT] OF ST_UpsDesiredSet;
	(* BMS 랙 선택표 (BMS 40001 랙 비트, 비트 n-1 = 랙 n). EMS 랙 명령(11·12)으로 바뀜. 0 = 저장 안 됨 → 설치된 랙 전부 *)
	g_awBmsRackMask	: ARRAY[1..GVL_PARAM.BMS_COUNT] OF WORD;

	(* 지령 거르기·시퀀스 (코어) *)
	g_stCmdFilter	: ST_CmdFilterSet := (
						bBadValue		:= TRUE,	fBadFactor	:= 1.5);	// 이상값: NaN·무한대 + 정격 × 1.5 초과 무시 (Auto·Manual)
	g_stManualCmdSet	: ST_ManualCmdSet := (
						bReverse		:= TRUE,	fDirBand	:= 1.0,	// Manual 방향 반대 지령 무시 (정격 1% 이하는 멈춘 것)
						bClearOnStop	:= TRUE);					// Manual: Run 확인 뒤 들어온 지령만 씀
	g_stSeqSet		: ST_SeqSet := (							// 시퀀스: 쓰기 주기, 명령 확인·재시도, 배터리 투입
						tWritePeriod	:= T#200MS,
						stPcs := (
							tCmdConfirm		:= T#30S,
							tStopRetry		:= T#5S,
							nStopRetry		:= 3,
							bStopRamp		:= FALSE,
							fStopDonePct	:= 1.0,
							tStopRampMax	:= T#30S),
						stBat := (
							eClose			:= E_BatClose.OnStart,
							bOpenOnStop		:= FALSE,
							tConfirm		:= T#60S,
							tOpenRetry		:= T#5S,
							nOpenRetry		:= 3));
	(* 현장 모듈 설정 (모듈마다 칸 하나, 타입 ST_ModuleSet은 90_Project). MAIN 액션 A_PassModuleSet에서 각 모듈 i_stSet에 넘김 *)
	g_stModuleSet	: ST_ModuleSet;

	(* MQTT 브로커 끊김 감시 [9번 수정 2026-11-09: 추가]. 고른 브로커 접속이 tLostDelay 넘게 끊기면 '브로커 끊김' 알람 + 운전 모드 요청을 모두 Manual로 (한 번, 다시 접속하면 다시 무장) *)
	g_stBrokerWatch	: ST_BrokerWatchSet;	// 기본: Local 브로커, 30 s

	(* 재기동 기록 (FB_AliveRecorder가 1 s마다 갱신, 파일 저장은 주기 저장) *)
	g_nLastAliveLocal	: ULINT;	// 마지막 동작 시각 (FILETIME 모양, 현지 시각). 2026-11-03 UTC(g_nLastAlive) → 현지로 바꾸며 이름 바꿈: 바꾼 뒤 첫 시작은 '기록 없음'
	g_sLastAlive	: STRING(31);	// 같은 시각, 현지 시각 글자
END_VAR

// ---- 90_Project/GVL_SITE.TcGVL
VAR_GLOBAL CONSTANT
	(* ================================================================
	   현장 구성 (현장이 바뀌면 재빌드)
	   ================================================================ *)
	(* UPS 연결: UPS 번호 1 → BMS 등록 칸 1 (현장 5: UPS 1대·BAT 1대). PCS 등록과는 별개.
	   UPS는 별도 I_Ups 드라이버이며 이 표는 UPS와 BMS의 소속 관계를 정의한다. *)
	UPS_BMS			: ARRAY[1..GVL_PARAM.UPS_COUNT] OF UINT := [1];

	(* 유닛 → PCS·배터리 그룹·제어 그룹 *)
	UNIT_CFG		: ARRAY[1..GVL_PARAM.UNIT_COUNT] OF ST_UnitCfg := [
						(nPcs := 1, nSub := 1, nBatGroup := 1, nGroup := 1, fPRated := 1000.0, fQRated := 500.0, fSRated := 1118.0),	// 유닛 1 = PCS1
						(nPcs := 2, nSub := 1, nBatGroup := 1, nGroup := 1, fPRated := 1000.0, fQRated := 500.0, fSRated := 1118.0)];	// 유닛 2 = PCS2 (배터리 그룹 2, 접속점은 유닛 1과 같음)
	(* BMS → 배터리 그룹. 유닛 n : BMS m = 같은 배터리 그룹 번호 *)
	BMS_CFG			: ARRAY[1..GVL_PARAM.BMS_COUNT] OF ST_BmsCfg := [
						(nBatGroup := 1, fCapacity := 0.0)];	// BMS 1 = 배터리 그룹 1 (UPS1 배터리). 용량 미정 (0 = SOC 균등)
	(* 계측점 = 계측기 값을 부호와 함께 더한 것 (계측기 값은 방전·공급 +)
	   예) Helios 기준점(VCB1): [(nMeter := 1, fSign := 1.0)]   CTPT 미터 (Beckhoff, PV 측)
	       Helios VCB2의 PV 값: [(nMeter := 1, fSign := 1.0), (nMeter := 2, fSign := -1.0)]   CTPT 미터 − ESS 미터
	       메시즈 수전점: [(nMeter := 1, fSign := -1.0)]   역전력계전기 (수전 +)를 뒤집음 *)
	POINT_CFG		: ARRAY[1..GVL_PARAM.POINT_COUNT] OF ST_PointCfg := [
						(astTerm := [(nMeter := 1, fSign := 1.0)])];	// 계측점 1 = 계측기 1
	GROUP_CFG		: ARRAY[1..GVL_PARAM.GROUP_COUNT] OF ST_GroupCfg := [
						(nPccPoint := 0)];	// no ESS PCC at this UPS-only site

	START_MODE		: ARRAY[1..GVL_PARAM.UNIT_COUNT] OF E_StartMode := [
						E_StartMode.Step, E_StartMode.Step];			// 유닛별 기동 방식

	(* MQTT 접속 (PRG_Mqtt → FB_MqttMain). 브로커 계정은 저장소에 올리지 않으려고 비워 둠: 빌드·다운로드 전에 sUserName·sUserPassword에 적고 이 두 줄은 커밋하지 않는다.
	   접속 값은 첫 호출 때 한 번 읽으므로 바꾸면 재빌드. 안 쓰는 브로커는 bUse := FALSE (지금은 PCS 값을 발행 직전 구조체까지만 시험하느라 모두 FALSE. 발행 시험 때 TRUE로) *)
	MQTT_SET		: ST_MqttSet := (
						nSiteId			:= 5,
						stCloud			:= (bUse := FALSE, sHost := '10.0.0.0', nPort := 1883),
						stLocal			:= (bUse := TRUE, sHost := '10.0.0.36', nPort := 1883),	// DGS MQTT 브로커 (현장 5). 브로커 끊김 감시 기본(Local)이 이 칸을 봄
						stAzure			:= (bUse := FALSE, sHost := '10.0.0.3', nPort := 1883),
						sUserName		:= 'dgs_admin',
						sUserPassword	:= '');

	(* 시험 모드: 사무실 가상 장비 시험용. 현장 빌드는 FALSE (가상 장비 연결 PRG_SimLink, 가상신호 GVL_TEST.g_astVirtual, 시험 리셋 GVL_TEST.g_bTestReset을 안 씀) *)
	TEST_MODE		: BOOL := FALSE; // real-map commissioning: no fabricated measurements

	(* 장비 쓰기 스위치: FALSE면 PMS는 계산·보고만 하고 PCS·BMS·보조 출력에 아무것도 쓰지 않음 (읽기 전용 시험).
	   실제 장비에 처음 연결할 때는 FALSE로 시작하고, 읽기 값이 맞는지 확인한 뒤 TRUE. 가상 장비 시험은 TRUE *)
	DEVICE_WRITE	: BOOL := FALSE;		// 제어 시험(PCS 시뮬레이터 192.168.0.120:602) 동안 TRUE. 실제 장비에 연결할 때는 FALSE로 시작

	(* 명령 필터·Manual 지령 거르기·시퀀스 설정은 운전 중 바꾸도록 GVL_PERSIST로 옮김 (g_stCmdFilter, g_stManualCmdSet, g_stSeqSet) *)

	(* 운전 모드 전환: 어디까지 하고 바꾸나 (Direct / Zero / Standby) *)
	MODE_SET		: ST_ModeSet := (
						eToManual		:= E_ModeSwitch.Standby,	// 출력 0 → 400 ms → Standby → 멈춤 확인 → Manual (Helios와 같음)
						eToAuto			:= E_ModeSwitch.Zero,		// 출력 0 → 400 ms → Auto
						tDelay			:= T#400MS,
						bKeepOnRestart	:= FALSE);	// PMS가 다시 켜지면 모든 유닛 Manual로 시작 (정전 뒤 장비 투입은 운전원이). TRUE = 저장된 모드 유지

	(* 이중화: 두 PLC에 같은 프로그램. 역할(Primary/Secondary)은 이 PLC의 AMS Net ID로 정함 (PRG_Redundancy)
	   이중화를 쓰면 bUse := TRUE, 두 PLC의 Net ID를 적음 (TwinCAT 시스템 화면 또는 온라인 PRG_Redundancy.sMyNetId) *)
	RED_SET			: ST_RedSet := (
						bUse			:= FALSE,
						sPrimaryNetId	:= '',
						sSecondaryNetId	:= '');

	(* 로그 설정 *)
	LOG_SET			: ST_LogSet := (
						tHold			:= T#10S,		// 출력 제한 이유가 이 시간 이상 유지될 때만 기록
						tPersistSave	:= T#60S,		// PERSISTENT 주기 저장 (설정 변경은 바로 저장)
						bUnitLimited	:= FALSE,		// 자세한 기록 (시운전·문제 추적 때 TRUE)
						bReqRefused		:= FALSE,
						bSeqChange		:= FALSE,
						bModeChange		:= FALSE,
						bBatRefused		:= TRUE,		// 배터리 요청 거부
						bCmdRefused		:= TRUE);		// 무시한 지령 (이상값·방향 반대)
END_VAR

VAR_GLOBAL

	(* ================================================================
	   장비·모듈 인스턴스
	   - 모듈 ID는 현장 안에서 겹치지 않게: 1~99 장비, 100~199 지령원, 200~ 기능 모듈
	   - 이름은 영문 (로그에 그대로 나옴)
	   - 장비 읽기 주기: 기본 200 ms. 장비마다 바꾸려면 선언에 추가 → (i_nModuleId := 1, i_sName := 'PCS1', i_tReadPeriod := T#500MS)
	   ================================================================ *)

	(* ---------- 장비: 기존 PCS 시험 인스턴스는 보관만 하며 g_aipPcs에는 등록하지 않는다 ---------- *)
	g_fbPcs1		: FB_PlaspoPcs	:= (i_nModuleId := 1, i_sName := 'PCS1', i_sIpAddr := '192.168.0.120', i_nPort := 602);
	g_fbPcs2		: FB_PcsSim		:= (i_nModuleId := 2, i_sName := 'PCS2');
	// 가상 PCS로 되돌리려면: g_fbPcs1 : FB_PcsSim := (i_nModuleId := 1, i_sName := 'PCS1');  (g_fbRptPcs1·MAIN A_Report의 RawMap 줄도 같이 뺌)
	// 보고 매핑 (PCS 1 → MQTT pcs 레코드). 배율은 플라스포 레지스터 맵 확인 후 i_f…Scale에 줌. MAIN 액션 A_Report가 부름
	g_fbRptPcs1		: FB_RptPlaspoPcs;
	// 실제 PCS 예: g_fbPcs1 : FB_PlaspoPcs := (i_nModuleId := 1, i_sName := 'PCS1', i_sIpAddr := '192.168.0.100', i_tReadPeriod := T#1S);
	g_fbBms1		: FB_EsolutionBms := (i_nModuleId := 11, i_sName := 'BMS1', i_nRackCount := GVL_PARAM.RACKS_PER_BMS, i_bReadDetails := TRUE, i_bEnable := TRUE, i_sIpAddr := '192.168.0.138', i_nPort := 504, i_nUnitId := 1); // 시험용: PC의 BMS 시뮬레이터 (03. simulator\ups_bms_sim.py)
	g_fbMeter1		: FB_MeterSim	:= (i_nModuleId := 21, i_sName := 'PCC1');

	(* UPS-only devices. TCP endpoints are deliberately empty and i_bEnable defaults FALSE.
	   Set each endpoint from the equipment list before read-only commissioning. *)
	g_fbUps1 : FB_SebangUps := (i_nModuleId := 41, i_sName := 'UPS1', i_bEnable := TRUE, i_sIpAddr := '192.168.0.138', i_nPort := 503, i_nUnitId := 1); // 시험용: PC의 UPS 시뮬레이터 (03. simulator\ups_bms_sim.py)
	g_aipUps : ARRAY[1..GVL_PARAM.UPS_COUNT] OF I_Ups := [g_fbUps1];	// 현장 5: UPS 1대

	(* ---------- 보조 장비: Helios에서 가져온 센서 드라이버 (2026-11-09). 맵·주소 미확보라 모두 i_bEnable FALSE (통신 안 함)
	   쓰려면 주소를 적고 i_bEnable := TRUE. 점 번호는 각 드라이버 머리 주석. 보호 판정은 아래 "보조 장비·규칙 예"처럼 FB_RuleBit·FB_RuleValue로 등록 ---------- *)
	g_fbThd1		: FB_AutonicsThd		:= (i_nModuleId := 32, i_sName := 'THD1', i_nSensorCount := 1, i_tReadPeriod := T#300MS);	// 오토닉스 온습도 (RTU, EL6022 채널). 채널 연결은 XAE I/O 화면에서. AI 1 온도·2 습도
	g_fbImd1		: FB_LsImd1000		:= (i_nModuleId := 33, i_sName := 'IMD1', i_tReadPeriod := T#1S);	// LS IMD1000 절연감시 (LS ETH-RSTP-DC24V 컨버터, 라벨 MAC 00-0B-29-00-6D-F7). 컨버터 IP 미확인이라 통신 끔: 라벨 초기값 192.168.0.100·종이 10.0.0.50 모두 응답 없음, 192.168.0.50은 다른 장비(ASUS). 찾으면 i_bEnable := TRUE, i_sIpAddr DI 1 경고·2 절연 경보, AI 1 절연저항. MAIN.A_Report가 q_stState로 imd 토픽 보고
	g_fbRio1		: FB_RootechAcuraIo	:= (i_nModuleId := 34, i_sName := 'RIO1');	// 루텍 ACURA3700 원격 I/O (TCP). i_sIpAddr 미정. DI 1..8 = 화재(열)·연기·가스 감지기 접점 (Helios 배치, 현장 결선 확인)
	g_fbThd2		: FB_ItGuardIeSx		:= (i_nModuleId := 35, i_sName := 'THD2', i_tReadPeriod := T#1S, i_bEnable := TRUE, i_sIpAddr := '192.168.0.70');	// ITGuard IE-SX 이더넷 온습도계 (TCP, 2026-11-09 PC에서 읽어 확인). AI 1 온도·2 습도. MAIN.A_Report가 temperature_sensor 토픽 보고
	g_fbGfr1		: FB_WoonyoungGfr	:= (i_nModuleId := 36, i_sName := 'GFR1', i_tReadPeriod := T#1S, i_nChannels := 8, i_nUnitId := 1, i_bEnable := TRUE);	// 운영 WYGF-D08NC 지락검출계전기 (RTU, EL6022 채널. _fbRtu InData·OutData를 XAE I/O에서 연결). AC 회로 누전. DI n 지락, AI n 누설전류 A
	g_fbAsd57		: FB_GasdnaAsd57		:= (i_nModuleId := 37, i_sName := 'ASD1', i_tReadPeriod := T#1S, i_nUnitId := 1, i_bEnable := TRUE);	// 가스디엔에이 ASD-57 열연복합 감지기 (RTU 9600 고정, EL6022 채널. 지락계전기와 다른 채널. _fbRtu InData·OutData를 XAE I/O에서 연결). DI 1 연기·2 온도 알람, AI 1·2 연기, 3 온도
	g_fbSmoke2		: FB_RuleBit			:= (i_nModuleId := 206, i_sName := 'Smoke2', i_ipAux := g_fbAsd57, i_nPoint := 1);	// 연기 감지 (ASD-57 연기 알람). 알람만 (조치 없음, 사고·고장 단계는 EMS). 2026-11-10
	g_fbIo1			: FB_AuxIo			:= (i_nModuleId := 31, i_sName := 'IO1');	// 벡호프 단자 I/O (EL1xxx DI). 점은 XAE I/O 화면에서 _abDi[n]에 연결. DI 1 = 가스디엔에이 TS-60 연기 접점 (흰 NO·초록 COM, 경보 때 닫힘). 2026-11-10
	g_fbSmoke1		: FB_RuleBit			:= (i_nModuleId := 205, i_sName := 'Smoke1', i_ipAux := g_fbIo1, i_nPoint := 1);	// 연기 감지 (TS-60 연기 접점). 알람만 (조치 없음, 사고·고장 단계는 EMS가 판단). 온도 접점(노랑·파랑)은 쓰지 않음 (사용자 2026-11-10)

	(* ---------- 지령원 ---------- *)
	g_fbSrcTest		: FB_SrcTest	:= (i_nModuleId := 101, i_sName := 'Test');
	(* ---------- 제어 모드: 접속점 그룹마다 관리자 하나 + 모드 한 세트 (접속점 그룹 안 Auto 유닛은 같은 모드). 모듈 ID 240~
	   [16번 수정 2026-11-09: PCS마다(유닛 단위) → 접속점 그룹 단위로 바꿈. 원래 g_fbCtrlMode1(유닛 1)·g_fbCtrlMode2(유닛 2)와 모드 두 세트 (ID 103, 244~247, 249)]
	   - 관리자 i_nUnit = 0: 접속점 그룹 하나를 통째로 맡음. 모드는 접속점 그룹 값(접속점·정격·SOC)을 보고 접속점 그룹 지령(접속점 기준)을 내고, 코어 분배가 접속점 그룹의 Auto 유닛에 나눔. Manual 유닛은 제어 모드를 받지 않음
	   - 스탠다드 스케줄(5)만 유닛별 값: EMS가 PCS마다 보낸 P를 그 PCS의 유닛에 그대로 냄 (ST_CtrlModeOut.bUnitOut)
	   - HMI가 관리자 i_nModeReq(모드 칸 번호, 0 = 없음)를 씀. 칸 번호 = g_aipCtrlMode1 순서. PERSISTENT가 아니라 재기동하면 0 (14번 탭 2번 결정)
	   - 설정은 GVL_PERSIST.g_stModuleSet 칸 (stCtrlMode1·stCmConstP1·stCmSchedule1·stCmPeakCut1·stCmSchedPeak1, 공통 stCmCommon)을 MAIN 액션 A_PassModuleSet에서 넘김. 피크 목표·정출력 값은 접속점 그룹 전체 값
	   - 접속점 그룹을 늘리면: 관리자·모드 5개 선언(등록 nGroup = 그 접속점 그룹) + 등록(g_aipSource·g_aipCtrlModeN·GVL_PERSIST.g_astSourceReg) + ST_ModuleSet 칸 + A_PassModuleSet 줄 + FB_ConfigCheck·FB_EventLog 입력 ---------- *)
	g_fbCtrlMode1	: FB_CtrlModeMgr	:= (i_nModuleId := 102, i_sName := 'CtrlMode1', i_nUnit := 0);	// 접속점 그룹 1 (접속점 그룹 단위). 설정 stCtrlMode1
	g_fbCmConstP1	: FB_CmConstPower	:= (i_nModuleId := 240, i_sName := 'CmConstP1');	// 1 정출력 (설정 stCmConstP1, 접속점 그룹의 접속점 기준 값)
	g_fbCmSchedule1	: FB_CmSchedule		:= (i_nModuleId := 241, i_sName := 'CmSchedule1');	// 2 스케줄 (시간표 stCmSchedule1, 접속점 그룹 값)
	g_fbCmPeakCut1	: FB_CmPeakCut		:= (i_nModuleId := 242, i_sName := 'CmPeakCut1');	// 3 피크컷 (설정 stCmPeakCut1, 목표 피크 = 접속점 그룹 전체)
	g_fbCmSchedPeak1	: FB_CmSchedPeak	:= (i_nModuleId := 243, i_sName := 'CmSchedPeak1');	// 4 통합 = 스케줄 + 피크컷 (시간표 stCmSchedule1, 설정 stCmSchedPeak1)
	g_fbCmStdSched1	: FB_CmStdSchedule	:= (i_nModuleId := 248, i_sName := 'CmStdSched1');	// 5 스탠다드 스케줄 = EMS 지령을 그대로 따름 (PCS마다 값, MAIN A_PassEmsCmd가 넘김)
	// EMS 지령원 (MQTT command). 상태 명령은 Auto에서 받고 충전·방전 P 지령은 i_bPEnable이 켜질 때만 냄. 입력은 MAIN 액션 A_PassEmsCmd가 넘김
	g_fbSrcEms		: FB_SrcEms		:= (i_nModuleId := 104, i_sName := 'Ems');

	(* ---------- SOC 정책 (버스 제한. 기본 등록: 모든 버스, Auto·Manual 모두. 적용 모드는 GVL_PERSIST.g_astBatRuleReg bAuto·bManual)
	   설정(한계·감발 폭·재개 마진)은 GVL_PERSIST.g_stModuleSet.stSocLimit, MAIN 액션 A_PassModuleSet에서 넘김 ---------- *)
	g_fbSocLimit	: FB_SocLimit	:= (i_nModuleId := 210, i_sName := 'SocLimit');	// SOC 감발·막음·재개 마진. 한도 0이면 그 방향 출력 0 (= 대기)

	(* ---------- 사용자 한도 (유닛 제한. EMS config pcs 충·방전 전력 한도도 여기에 씀: FB_EmsConfigApply) [9-21 수정 2026-11-04: 아래 주석 예에서 꺼내 기본 등록.
	   설정 stUnitLimit 기본 모두 끔 → 켜기 전에는 하는 일 없음. 적용 모드는 GVL_PERSIST.g_astUnitRuleReg[1] (기본 전체 유닛, Auto·Manual)] ---------- *)
	g_fbUnitLimit	: FB_UnitLimit := (i_nModuleId := 230, i_sName := 'UserLimit');	// 설정 stUnitLimit

	(* ---------- 표준 보호 (기본 등록. 빼면 그 보호 없음. 설정은 GVL_PERSIST.g_astRuleCfg 같은 칸) ---------- *)
	g_fbProtPcsFault	: FB_ProtPcsFault	:= (i_nModuleId := 901, i_sName := 'PcsFault');
	g_fbProtPcsComm		: FB_ProtPcsComm	:= (i_nModuleId := 902, i_sName := 'PcsComm');
	g_fbProtBmsFault	: FB_ProtBmsFault	:= (i_nModuleId := 903, i_sName := 'BmsFault');
	g_fbProtBmsComm		: FB_ProtBmsComm	:= (i_nModuleId := 904, i_sName := 'BmsComm');
	g_fbProtPccInvalid	: FB_ProtPccInvalid	:= (i_nModuleId := 905, i_sName := 'PccInvalid');
	g_fbProtRespStd		: FB_ProtRespStd		:= (i_nModuleId := 900, i_sName := 'RespStd');	// 표준 대응: 칸 설정(g_astRuleCfg.stProt)의 조치. 칸마다 같은 인스턴스

	(* ---------- 보조 장비·규칙 예 (현장에서 주석을 풀어 씀)
	Helios 센서로 쓰는 예 (위 g_fbThd1·g_fbImd1·g_fbRio1):
	g_fbFireHeat	: FB_RuleBit	:= (i_nModuleId := 204, i_sName := 'FireHeat', i_ipAux := g_fbRio1, i_nPoint := 1);	// 화재(열) 감지기 접점
	g_fbFireSmoke	: FB_RuleBit	:= (i_nModuleId := 205, i_sName := 'FireSmoke', i_ipAux := g_fbRio1, i_nPoint := 2);	// 연기 감지기 접점
	g_fbFireGas		: FB_RuleBit	:= (i_nModuleId := 206, i_sName := 'FireGas', i_ipAux := g_fbRio1, i_nPoint := 3);	// 가스 감지기 접점
	g_fbImdFault	: FB_RuleBit	:= (i_nModuleId := 207, i_sName := 'ImdFault', i_ipAux := g_fbImd1, i_nPoint := 2);	// IMD 고장 (경고까지 보려면 점 1도 한 칸 더)
	g_fbRoomTemp	: FB_RuleValue	:= (i_nModuleId := 208, i_sName := 'RoomTemp', i_ipAux := g_fbThd1, i_nPoint := 1);	// 실내 온도
	등록은 아래 g_fbFire 예와 같음 (g_aipRule 칸 + RULE_COUNT + GVL_PERSIST.g_astRuleCfg 같은 칸, 대응을 비우면 알람만)
	g_fbIo1			: FB_AuxIo		:= (i_nModuleId := 31, i_sName := 'IO1', i_afAiGain := [0.1, 0.1]);		// 점은 화면에서 연결
	g_fbFire		: FB_RuleBit	:= (i_nModuleId := 201, i_sName := 'Fire', i_ipAux := g_fbIo1, i_nPoint := 1);			// 설정 stFire
	g_fbEStop		: FB_RuleBit	:= (i_nModuleId := 202, i_sName := 'EStopSw', i_ipAux := g_fbIo1, i_nPoint := 2);		// 설정 stEStop (b접점, 통신 끊김 시 조건)
	g_fbBatTemp		: FB_RuleValue	:= (i_nModuleId := 203, i_sName := 'BatRoomTemp', i_ipAux := g_fbIo1, i_nPoint := 1);	// 설정 stBatTemp (해소 폭 2.0)
	등록: g_aipAux := [g_fbIo1], g_aipRule := [표준 5개, g_fbFire, g_fbEStop, g_fbBatTemp] (보호 6~8칸, RULE_COUNT 8), g_aipOutput := [g_fbBatTemp] (팬 켜기)
	      같은 규칙을 보호와 출력에 함께 등록할 수 있음. 설정은 GVL_PERSIST.g_astRuleCfg / g_astOutputCfg 같은 칸 번호
	      모듈 설정(b접점·해소 폭 등)은 GVL_PERSIST.g_stModuleSet 칸 + MAIN 액션 A_PassModuleSet
	차단기(VCB) 운전원 투입·개방 예:
	g_fbVcb1		: FB_BreakerCtrl := (i_nModuleId := 220, i_sName := 'VCB1', i_ipAux := g_fbIo1, i_nClosedPoint := 3);	// 상태 접점 DI 3, 설정 stVcb1
	등록: g_aipOutput 두 칸에 g_fbVcb1 (g_astOutputCfg: 투입 코일 칸 fThreshold := 1, 개방 코일 칸 fThreshold := 2, nAux·nPoint = 코일 DO, 지연 0·유지 끔),
	      g_aipRule 한 칸에 g_fbVcb1 (g_astRuleCfg: 조치 None = 투입·개방 실패 알람만). HMI는 g_fbVcb1.i_bCloseCmd·i_bOpenCmd·i_bResetFail을 켬
	사용자 한도 (유닛마다 P·Q 상·하한 kW·kvar) 예:
	(9-21 수정 2026-11-04: 위 SOC 정책 다음으로 꺼내 기본 등록함) g_fbUnitLimit	: FB_UnitLimit := (i_nModuleId := 230, i_sName := 'UserLimit');	// 설정 stUnitLimit
	등록: g_aipUnitRule 한 칸에 g_fbUnitLimit (g_astUnitRuleReg: nTarget 0 = 전체 유닛, bAuto·bManual로 적용 모드)
	---------- *)

	(* ================================================================
	   등록 (선언할 때 연결. 다른 곳에서 쓰지 않음)
	   - 칸을 비워 두면 그 기능은 없다
	   ================================================================ *)
	g_aipPcs		: ARRAY[1..GVL_PARAM.PCS_COUNT] OF I_Pcs; // UPS site: no separate PCS installed
	g_aipBms		: ARRAY[1..GVL_PARAM.BMS_COUNT] OF I_Bms				:= [g_fbBms1];	// 현장 5: BAT 1대
	g_aipMeter		: ARRAY[1..GVL_PARAM.METER_COUNT] OF I_Meter; // no separate PCC meter in UPS-only commissioning
	g_aipAux		: ARRAY[1..GVL_PARAM.AUX_COUNT] OF I_AuxDevice		:= [g_fbThd1, g_fbImd1, g_fbRio1, g_fbThd2, g_fbGfr1, g_fbIo1, g_fbAsd57];	// 보조 장비 (규칙·출력 설정의 nAux = 칸 번호)
	g_aipSource		: ARRAY[1..GVL_PARAM.SOURCE_COUNT] OF I_CommandSource; // ESS command sources unregistered at UPS site	// 등록표 GVL_PERSIST.g_astSourceReg 같은 칸
	g_aipLimit		: ARRAY[1..GVL_PARAM.LIMIT_COUNT] OF I_LimitRule;
	g_aipPermit		: ARRAY[1..GVL_PARAM.PERMIT_COUNT] OF I_StartPermit;
	g_aipComp		: ARRAY[1..GVL_PARAM.COMP_COUNT] OF I_Compensator;
	g_aipRule		: ARRAY[1..GVL_PARAM.RULE_COUNT] OF I_ProtectionRule	:= [g_fbProtPcsFault, g_fbProtPcsComm, g_fbProtBmsFault, g_fbProtBmsComm, g_fbProtPccInvalid, g_fbSmoke1, g_fbSmoke2];	// 보호 (설정 g_astRuleCfg). 1~5 = 표준 보호, 6 = 연기 TS-60, 7 = 연기 ASD-57 (대응 칸 비움 = 알람만)
	g_aipResp		: ARRAY[1..GVL_PARAM.RULE_COUNT] OF I_ProtResponse	:= [g_fbProtRespStd, g_fbProtRespStd, g_fbProtRespStd, g_fbProtRespStd, g_fbProtRespStd];	// 보호 대응 (같은 칸). 1~5 = 표준 대응. 비우면 조치 없음 (알람만). 현장 보호 칸을 늘리면 그 칸에도 등록
	g_aipOutput	: ARRAY[1..GVL_PARAM.OUTPUT_COUNT] OF I_OutputRule;	// 보조 장비 출력 규칙
	g_aipUnitRule	: ARRAY[1..GVL_PARAM.UNIT_RULE_COUNT] OF I_UnitLimitRule	:= [g_fbUnitLimit];	// 유닛 제한 (등록 설정 GVL_PERSIST.g_astUnitRuleReg). 1 = 사용자 한도 [9-21 수정 2026-11-04: 등록. 원래 빈 칸]
	g_aipBatRule	: ARRAY[1..GVL_PARAM.BAT_RULE_COUNT] OF I_BatLimitRule	:= [g_fbSocLimit];	// 버스 제한 (g_astBatRuleReg). 1 = SOC 정책
	g_aipCtrlMode1		: ARRAY[1..GVL_PARAM.CTRL_MODE_COUNT] OF I_ControlMode	:= [g_fbCmConstP1, g_fbCmSchedule1, g_fbCmPeakCut1, g_fbCmSchedPeak1, g_fbCmStdSched1];	// 접속점 그룹 1 제어 모드 (칸 번호 = g_fbCtrlMode1.i_nModeReq). MAIN A_PassModuleSet이 관리자에 넘김 [16번 수정 2026-11-09: g_aipCtrlMode2 없앰]
	g_aipSelectPolicy	: ARRAY[1..GVL_PARAM.GROUP_COUNT] OF I_SelectPolicy;	// 그룹별 지령원 고르기 정책. 비우면 코어 기본 (g_astGroupSet eSelP·eSelQ)
	g_aipDistPolicy		: ARRAY[1..GVL_PARAM.GROUP_COUNT] OF I_DistPolicy;		// 그룹별 분배 정책. 비우면 코어 기본 (g_astGroupSet eDistBasis)
	g_ipAutoGate		: I_Gate;		// Auto 지령 거르기. 비우면 코어 기본 (통과)
	g_ipManualGate		: I_Gate;		// Manual 지령 거르기. 비우면 코어 기본 (방향 반대 무시·Run 뒤 새 지령 대기, g_stManualCmdSet)
END_VAR

// ---- 90_Project/GVL_IF.TcGVL
VAR_GLOBAL
	g_nUpsConfigSeq : UDINT; // MqttTask writer, PlcTask reader; odd=in progress
	g_stUpsConfigRx : ST_IfUpsConfigRx;
	g_nUpsCmdSeq : UDINT; // UPS 명령 칸 번호. PRG_Mqtt(MqttTask)가 쓰고 MAIN(PlcTask)이 읽음. 홀수 = 쓰는 중
	g_astUpsCmd : ARRAY[1..GVL_PARAM.UPS_COUNT] OF ST_IfUpsCmd; // UPS별 마지막 명령 (번호가 바뀌면 새 명령)
	(* ================================================================
	   태스크 사이에 주고받는 값 (자리만. 내용은 인터페이스가 정해지면 채움)

	   규칙
	   - 칸마다 쓰는 태스크는 하나. 다른 태스크는 읽기만
	   - 쓰는 쪽: 쓰기 전에 번호(…Seq)를 1 올리고(홀수 = 쓰는 중), 내용을 다 쓴 뒤 다시 1 올림(짝수 = 끝)
	   - 읽는 쪽: 번호 읽기(짝수일 때만) → 내용 복사 → 번호 다시 읽기. 두 번호가 같을 때만 새 값으로 씀
	     (쓰는 도중에 읽어 반만 바뀐 값을 쓰지 않게. 우선순위가 높은 태스크가 쓰는 중에 끼어들어도 읽는 쪽이 걸러냄.
	      내용 쪽에도 …RxCount·nSeq 같은 번호를 두어 새 값인지는 그 번호로 가림)
	   - 제어 흐름(읽기 → 보호 → 요청 → 중재 → 분배 → 쓰기)은 PlcTask의 MAIN에만 둔다
	   - 태스크 전용 FB 인스턴스는 그 태스크 PRG 안에 선언한다. I/O 연결이 있는 인스턴스를 GVL에 두면
	     {attribute 'TcContextName' := '태스크 이름'}을 붙여야 그 태스크 주기로 I/O가 갱신된다 (기본은 PlcTask)
	   ================================================================ *)

	(* ---------- MAIN → MQTT: 보고 (쓰는 곳: MAIN의 FB_Report) ---------- *)
	g_nReportSeq		: UDINT;		// 보고 칸 번호 (홀수 = 쓰는 중, 짝수 = 끝). MAIN 액션 A_Report가 씀
	g_stReport			: ST_IfReport;	// 발행 직전 PCS 레코드 (보고 매핑 모듈 결과). PRG_Mqtt가 복사해 GVL_MQTT.g_stPcsPublish에 채움

	(* ---------- MQTT → MAIN: 명령 (쓰는 곳: PRG_Mqtt) ---------- *)
	g_nCmdSeq			: UDINT;		// 명령 칸 번호 (홀수 = 쓰는 중, 짝수 = 끝). PRG_Mqtt가 씀
	g_stEmsCmd			: ST_IfEmsCmd;	// EMS 명령: PCS·BMS 상태 명령과 충전·방전 P. PRG_Mqtt(FB_EmsCommand 결과)가 씀. MAIN 액션 A_PassEmsCmd가 복사해 지령원 FB_SrcEms에 넘김
	(* ---------- MQTT → MAIN: EMS config (쓰는 곳: PRG_Mqtt) [9-21 수정 2026-11-04: 추가] ---------- *)
	g_nCfgSeq			: UDINT;		// config 칸 번호 (홀수 = 쓰는 중, 짝수 = 끝). PRG_Mqtt가 씀
	g_stEmsCfg			: ST_IfEmsCfg;	// 받은 config 레코드(pcs·bat) + 칸마다 번호. MAIN 액션 A_PassEmsCfg가 복사해 FB_EmsConfigApply에 넘김
	(* ---------- MAIN → MQTT: config echo (쓰는 곳: MAIN) [9-21 수정 2026-11-04: 추가] ---------- *)
	g_nCfgEchoSeq		: UDINT;		// echo 칸 번호 (홀수 = 쓰는 중, 짝수 = 끝)
	g_stEmsCfgEcho		: ST_IfEmsCfgEcho;	// 실제 설정 (설정 보호 뒤). PRG_Mqtt가 복사해 config echo로 발행

	(* ---------- MQTT → MAIN: 브로커 접속 상태 (쓰는 곳: PRG_Mqtt) [9번 수정 2026-11-09: 추가]. 칸 1 Cloud, 2 Local, 3 Azure ---------- *)
	g_abBrokerUse		: ARRAY[1..3] OF BOOL;	// 쓰는 브로커 (GVL_SITE.MQTT_SET bUse)
	g_abBrokerConn		: ARRAY[1..3] OF BOOL;	// 구독 클라이언트가 브로커에 접속됨 (command·config를 받는 쪽)

	(* ---------- 빠른 계측 → MAIN (쓰는 곳: PRG_Fast) ---------- *)
	g_nFastSeq			: UDINT;		// 계측값을 다 쓴 뒤 올림. MAIN 쪽 계측기 드라이버가 읽음
	// 계측값 자리

	(* ---------- 이중화 (쓰는 곳: PRG_Redundancy) ---------- *)
	g_eRedRole			: E_RedRole;	// 이 PLC의 역할 (Primary/Secondary). 이중화를 안 쓰면 Primary
	g_bRedActive		: BOOL := NOT GVL_SITE.RED_SET.bUse;	// 이 PLC가 지금 장비에 쓰는가 (Active). 이중화를 안 쓰면 항상 TRUE, 쓰면 역할이 정해질 때까지 FALSE
	g_nRedSeq			: UDINT;		// 보낸 하트비트 수 (FB_RedLink)
	g_ePeerState		: E_RedPeer;	// 상대 PLC 상태 (EAP 하트비트 + 접점). 이중화를 안 쓰면 Unknown
	g_bPeerEapOk		: BOOL;			// EAP 하트비트 정상
	g_bPeerWireOk		: BOOL;			// 접점(alive) 신호 정상
	g_nPeerRole			: INT;			// 상대가 보낸 역할 (E_RedRole). EAP 정상일 때만 유효
	g_bPeerActive		: BOOL;			// 상대가 보낸 Active (EAP)
	g_bPeerWireActive	: BOOL;			// 상대 Active 접점 (EAP와 따로 봄)
	g_eRedState			: E_RedState;	// 이 PLC의 이중화 상태 (Init/Standby/Active/Failed). g_bRedActive는 이 상태가 Active인 것
	g_bRedRoleConflict	: BOOL;			// 두 PLC가 같은 역할 (설정 오류)
	g_bRedWrite			: BOOL := NOT GVL_SITE.RED_SET.bUse;	// 장비에 써도 됨 = Active가 된 뒤 tWriteHold 지남 (MAIN의 bWriteEnable이 봄). 이중화를 안 쓰면 항상 TRUE
	g_nPeerState		: INT;			// 상대가 보낸 이중화 상태 (E_RedState). EAP 정상일 때만 유효
	g_bSyncInSync		: BOOL;			// 상대 Active의 설정과 내 설정이 같음 (내가 Active가 아닐 때만 TRUE). 복귀 조건
	g_bSyncFresh		: BOOL;			// 상대가 보낸 동기화 값이 낡지 않음
	g_nSyncApplied		: UDINT;		// 상대 값으로 내 설정 블록을 덮어쓴 횟수
	g_nRedResumeCount	: UDINT;		// PLC가 멈췄다 이어진 횟수 (이 때 이중화 상태를 Init부터 다시 정함)
	g_nRedSwitchCount	: UDINT;		// Active가 바뀐 횟수 (들어가거나 나옴)
	g_eRedSwitch		: E_RedSwitch;	// Active가 바뀐 마지막 이유 (None/Start/PeerLost/Failback/Yield)
	// 동기화할 값 자리
END_VAR

// ---- 10_Core/01_Interface/I_UnitLimitRule.TcIO
INTERFACE I_UnitLimitRule EXTENDS I_Module

METHOD M_Evaluate : ST_LimitOut	// 유닛 P·Q 한도 (사용자 한도 등). bActive = FALSE면 제한 없음. 범위를 좁히기만 함 (0은 항상 허용)
VAR_INPUT
	i_stView	: ST_UnitLimitView;
END_VAR
END_METHOD

END_INTERFACE

// ---- 10_Core/01_Interface/I_BatLimitRule.TcIO
INTERFACE I_BatLimitRule EXTENDS I_Module

METHOD M_Evaluate : ST_BatLimitOut	// 배터리 버스 충·방전 한도 (SOC 감발 등). 범위를 좁히기만 함 (0은 항상 허용)
VAR_INPUT
	i_stView	: ST_BatLimitView;
END_VAR
END_METHOD

END_INTERFACE

// ---- 10_Core/01_Interface/I_Gate.TcIO
INTERFACE I_Gate EXTENDS I_Module	// 지령 거르기 (접수·보류·무시·새 지령 대기). 경로마다 한 칸 (GVL_SITE.g_ipAutoGate·g_ipManualGate), 비우면 코어 기본

METHOD M_Filter		// 매 스캔 한 번 (경로마다). 상태(보류 등)를 가져도 됨
VAR_INPUT
	i_stView	: ST_GateView;
END_VAR
VAR_IN_OUT CONSTANT
	iq_astUnitP		: ARRAY[1..GVL_PARAM.UNIT_COUNT] OF ST_Pick;		// 이 경로 FB_Select 결과 (다른 경로 유닛은 비활성)
	iq_astUnitQ		: ARRAY[1..GVL_PARAM.UNIT_COUNT] OF ST_Pick;
	iq_astGrpP		: ARRAY[1..GVL_PARAM.GROUP_COUNT] OF ST_Pick;
	iq_astGrpQ		: ARRAY[1..GVL_PARAM.GROUP_COUNT] OF ST_Pick;
	iq_aeOpMode		: ARRAY[1..GVL_PARAM.UNIT_COUNT] OF E_OpMode;		// 유닛 실제 운전 모드
	iq_astUnit		: ARRAY[1..GVL_PARAM.UNIT_COUNT] OF ST_UnitState;	// 유닛 상태 (실제 출력 방향·운전 상태)
	iq_astUnitCfg	: ARRAY[1..GVL_PARAM.UNIT_COUNT] OF ST_UnitCfg;
END_VAR
VAR_IN_OUT
	iq_stOut		: ST_GateOut;		// 거른 결과 (Gate가 채움. 지난 스캔 값이 남아 있음)
END_VAR
END_METHOD

END_INTERFACE

// ---- 10_Core/01_Interface/I_SelectPolicy.TcIO
INTERFACE I_SelectPolicy EXTENDS I_Module	// 고르기 정책: 지령원 후보 중 값 하나를 정함 (고르기·합치기). 그룹마다 한 칸 (GVL_SITE.g_aipSelectPolicy), 비우면 코어 기본 FB_SelectStd

METHOD M_Select : ST_Pick		// 고른 값. bActive = FALSE면 값 없음. 같은 입력이면 같은 결과 (한 스캔에 여러 번 부름, 상태를 바꾸지 않음)
VAR_INPUT
	i_stView	: ST_SelectView;
END_VAR
END_METHOD

END_INTERFACE

// ---- 10_Core/01_Interface/I_DistPolicy.TcIO
INTERFACE I_DistPolicy EXTENDS I_Module	// 분배 정책: 그룹 몫을 유닛에 나눌 무게. 그룹마다 한 칸 (GVL_SITE.g_aipDistPolicy), 비우면 코어 기본 FB_DistStd

METHOD M_Weight : REAL		// 이 유닛의 무게 (0 이상, 클수록 많이). 0 = 이 유닛에 안 줌. 같은 입력이면 같은 결과 (한 스캔에 여러 번 부름)
VAR_INPUT
	i_stView	: ST_DistView;
END_VAR
END_METHOD

END_INTERFACE

// ---- 10_Core/01_Interface/I_AuxDevice.TcIO
INTERFACE I_AuxDevice EXTENDS I_Module

METHOD M_Cycle
END_METHOD

PROPERTY Comm : BOOL
GET
END_GET
END_PROPERTY

METHOD M_GetValue : ST_Val
VAR_INPUT
	i_nPoint	: UINT;			// 장비 안의 아날로그 입력 점 번호
END_VAR
END_METHOD

METHOD M_GetBit : BOOL
VAR_INPUT
	i_nPoint	: UINT;			// 장비 안의 디지털 입력 점 번호
END_VAR
END_METHOD

METHOD M_SetBit		// 디지털 출력 점에 씀 (FB_AuxOutput만 부름)
VAR_INPUT
	i_nPoint	: UINT;			// 장비 안의 디지털 출력 점 번호
	i_bValue	: BOOL;
END_VAR
END_METHOD

METHOD M_SetValue		// 아날로그 출력 점에 씀
VAR_INPUT
	i_nPoint	: UINT;			// 장비 안의 아날로그 출력 점 번호
	i_fValue	: REAL;
END_VAR
END_METHOD

END_INTERFACE

// ---- 10_Core/01_Interface/I_OutputRule.TcIO
INTERFACE I_OutputRule EXTENDS I_Module		// 출력 규칙: 보조 장비 출력(DO)을 켤지 판단만. 쓰는 건 코어 FB_AuxOutput

METHOD M_Check : BOOL		// TRUE = 출력 켬 (지연·유지는 코어가 처리)
VAR_INPUT
	i_fThreshold	: REAL;			// ST_OutputCfg.fThreshold
END_VAR
END_METHOD

END_INTERFACE

// ---- 10_Core/01_Interface/I_Bms.TcIO
INTERFACE I_Bms EXTENDS I_Module

METHOD M_Cycle
END_METHOD

PROPERTY BatState : ST_BatState
GET
END_GET
END_PROPERTY

METHOD M_SetStateCmd : BOOL
VAR_INPUT
	i_stCmd		: ST_BatCmd;	// Close / Open / EStop / Reset
END_VAR
END_METHOD

END_INTERFACE

// ---- 10_Core/01_Interface/I_CommandSource.TcIO
INTERFACE I_CommandSource EXTENDS I_Module

METHOD M_Cycle
VAR_INPUT
	i_stReg		: ST_SourceReg;		// 등록표 한 줄
	i_stView	: ST_GroupView;		// 대상 그룹 값 (대상이 모든 그룹이면 그룹 1)
END_VAR
END_METHOD

PROPERTY Output : ST_SourceOutput
GET
END_GET
END_PROPERTY

END_INTERFACE

// ---- 10_Core/01_Interface/I_Compensator.TcIO
INTERFACE I_Compensator EXTENDS I_Module

METHOD M_Calc : ST_PQ			// 목표에 더할 보정량
VAR_INPUT
	i_stView	: ST_GroupView;
END_VAR
END_METHOD

END_INTERFACE

// ---- 10_Core/01_Interface/I_LimitRule.TcIO
INTERFACE I_LimitRule EXTENDS I_Module

PROPERTY Basis : E_LimitBasis
GET
END_GET
END_PROPERTY

METHOD M_Evaluate : ST_LimitOut
VAR_INPUT
	i_stView	: ST_GroupView;
END_VAR
END_METHOD

END_INTERFACE

// ---- 10_Core/01_Interface/I_Meter.TcIO
INTERFACE I_Meter EXTENDS I_Module

METHOD M_Cycle
END_METHOD

PROPERTY MeterState : ST_MeterState
GET
END_GET
END_PROPERTY

END_INTERFACE

// ---- 10_Core/01_Interface/I_Module.TcIO
INTERFACE I_Module EXTENDS __SYSTEM.IQueryInterface		// 모든 모듈의 공통. IQueryInterface: 같은 인스턴스인지 주소로 비교 (FB_ModuleList, __QUERYPOINTER)

PROPERTY ModuleId : UINT
GET
END_GET
END_PROPERTY

PROPERTY ModuleName : STRING(31)
GET
END_GET
END_PROPERTY

METHOD M_ReasonText : WSTRING(63)		// 이 모듈의 이유 코드 → 문구 (로그용)
VAR_INPUT
	i_nReason	: UINT;
END_VAR
END_METHOD

METHOD M_CheckSet : WSTRING(63)		// 이 모듈 설정 값 점검 (운전 중 HMI로 바꾸는 값). 빈 문구 = 정상, 아니면 오류 문구 (짧게) → FB_ConfigCheck가 설정 오류로 올림
END_METHOD

END_INTERFACE

// ---- 10_Core/01_Interface/I_Pcs.TcIO
INTERFACE I_Pcs EXTENDS I_Module

METHOD M_Cycle
END_METHOD

METHOD M_GetUnitState : ST_UnitState
VAR_INPUT
	i_nSub		: UINT;			// PCS 안의 유닛 번호
END_VAR
END_METHOD

METHOD M_SetPower : BOOL
VAR_INPUT
	i_nSub		: UINT;
	i_fP		: REAL;			// kW, 방전 +
	i_fQ		: REAL;			// kvar, 공급 +
END_VAR
END_METHOD

METHOD M_SetStateCmd : BOOL
VAR_INPUT
	i_nSub		: UINT;
	i_stCmd		: ST_PcsCmd;
END_VAR
END_METHOD

END_INTERFACE

// ---- 10_Core/01_Interface/I_ReqDevice.TcIO
INTERFACE I_ReqDevice EXTENDS I_Module		// 요청을 받는 새 장비 종류 (PCS·BMS·DO가 아닌 장비. 모양만 정함: 등록·코어 연결은 장비가 생길 때)
// 코어는 명령 내용을 모름: 장비마다 요청을 모아 센 쪽(M_CmdRank) 하나를 M_Request로 넘기고 요청 주체를 남김
// 장비 쓰기는 이 장비 모듈 한 곳 (R2: 장비 종류마다 한 곳). 장비 사이 순서(예: PCS 정지 확인 뒤 차단기 개방)는 보호 대응이 상태를 보고 진행

METHOD M_CmdRank : INT		// 명령 세기 (클수록 셈. 0 이하 = 요청 없음). 같은 장비에 요청이 겹치면 코어가 센 쪽 하나를 고름
VAR_INPUT
	i_nCmd		: UINT;		// 이 장비 모듈이 정한 명령 코드 (0 = 요청 없음)
END_VAR
END_METHOD

METHOD M_Request		// 코어가 합친 이번 스캔 요청 하나를 넘김 (요청 없으면 0). 명령·확인·재시도·실패 판단과 장비 쓰기는 장비 모듈이 함
VAR_INPUT
	i_nCmd		: UINT;		// 명령 코드 (0 = 요청 없음)
	i_nOrigin	: UINT;		// 요청한 모듈 ID (기록용)
END_VAR
END_METHOD

END_INTERFACE

// ---- 10_Core/01_Interface/I_ProtResponse.TcIO
INTERFACE I_ProtResponse EXTENDS I_Module		// 보호 대응: 조건이 걸리면 무엇을, 누구에게, 어떤 순서로 요청할지. 칸을 비우면 표준 대응 (FB_ProtRespStd, ST_ProtCfg)

METHOD M_Respond		// 보호 칸 하나·대상 하나의 대응: 무엇을, 누구에게 요청할지 iq_stReq에 씀. 장비에 직접 쓰지 않음
// 코어가 매 스캔 범위 안 대상마다 부름 (조건이 없을 때도: 단계 대응의 타이머·상태를 풀 수 있게). 대상 번호가 0으로 등록되면 대상마다 상태를 따로 둠
VAR_INPUT
	i_bActive		: BOOL;			// 보호 조건 있음 (등록 bAuto·bManual 중 하나가 켜져 있고 조건 모듈이 TRUE)
	i_tActive		: TIME;			// 조건이 이어진 시간 (조건 없으면 0)
	i_nTarget		: UINT;			// 대상 번호 (범위는 i_stRule.eScope. Site면 1)
	i_stRule		: ST_RuleCfg;		// 이 칸 설정 (범위·대상·임계값·표준 대응 설정)
END_VAR
VAR_IN_OUT CONSTANT
	iq_astUnit		: ARRAY[1..GVL_PARAM.UNIT_COUNT] OF ST_UnitState;	// 장비 상태 (이번 스캔 스냅샷, 읽기 전용)
	iq_astBms		: ARRAY[1..GVL_PARAM.BMS_COUNT] OF ST_BatState;
	iq_astUnitCfg	: ARRAY[1..GVL_PARAM.UNIT_COUNT] OF ST_UnitCfg;		// 소속 (제어 그룹·배터리 그룹)
	iq_astBmsCfg	: ARRAY[1..GVL_PARAM.BMS_COUNT] OF ST_BmsCfg;
	iq_aeOpMode		: ARRAY[1..GVL_PARAM.UNIT_COUNT] OF E_OpMode;		// 실제 운전 모드
END_VAR
VAR_IN_OUT
	iq_stReq		: ST_ProtReq;		// 요청 (코어가 비워서 넘김)
END_VAR
END_METHOD

END_INTERFACE

// ---- 10_Core/01_Interface/I_ProtectionRule.TcIO
INTERFACE I_ProtectionRule EXTENDS I_Module

METHOD M_Evaluate : BOOL		// TRUE = 보호 조건 있음. 판단만 함 (조치는 같은 칸의 대응, 비우면 표준 대응. 지연은 없음: 떨림 방지가 필요하면 모듈 설정에). 대상 번호가 0이면 코어가 범위 안 대상마다 한 번씩 부름
VAR_INPUT
	i_stView	: ST_ProtView;	// 대상 하나의 정보 (범위·대상 번호·임계값·상태)
END_VAR
END_METHOD

END_INTERFACE

// ---- 10_Core/01_Interface/I_StartPermit.TcIO
INTERFACE I_StartPermit EXTENDS I_Module

METHOD M_Evaluate : BOOL		// TRUE = 기동 허가
VAR_INPUT
	i_stView	: ST_GroupView;
	i_bRequest	: BOOL;				// 그룹이 기동을 기다리는 중
END_VAR
END_METHOD

PROPERTY Reason : UINT			// 허가하지 않은 이유 코드. 0 = 없음
GET
END_GET
END_PROPERTY

END_INTERFACE

// ---- 10_Core/01_Interface/I_ControlMode.TcIO
INTERFACE I_ControlMode EXTENDS I_Module	// 제어 모드 하나 (피크 저감·FR·스케줄·정출력 등). FB_CtrlModeMgr가 한 번에 하나만 켬. 켜진 동안에만 M_Calc를 부름

METHOD M_CheckEnter : UINT		// 지금 진입해도 되나. 0 = 됨, 그 외 = 이유 코드 (M_ReasonText). 상태를 바꾸지 않음 (한 스캔에 여러 번 부를 수 있음)
VAR_INPUT
	i_stView	: ST_CtrlModeView;	// 그룹 값(stGroup)·현지 시각(stTime). 관리자가 매 스캔 채움
END_VAR
END_METHOD

METHOD M_Enter		// 켜질 때 한 번. 내부 상태(타이머·적분 등) 초기화
VAR_INPUT
	i_stView	: ST_CtrlModeView;	// 그룹 값(stGroup)·현지 시각(stTime). 관리자가 매 스캔 채움
END_VAR
END_METHOD

METHOD M_Calc : ST_CtrlModeOut		// 켜져 있는 동안 매 스캔 한 번. 스스로 끝낼 때(bExitReq)도 그 스캔의 P·Q는 그대로 냄 (관리자가 0으로 넘김)
VAR_INPUT
	i_stView	: ST_CtrlModeView;	// 그룹 값(stGroup)·현지 시각(stTime). 관리자가 매 스캔 채움
END_VAR
END_METHOD

METHOD M_Exit		// 꺼질 때 한 번 (요청으로 바뀌든 스스로 끝내든)
END_METHOD

END_INTERFACE

// ---- 20_Module/Ups/I_Ups.TcIO
INTERFACE I_Ups EXTENDS I_Module

METHOD M_Cycle
END_METHOD

PROPERTY UpsState : ST_UpsState
GET
END_GET
END_PROPERTY

METHOD M_RequestCommand : BOOL
VAR_INPUT i_eCommand : E_UpsCommand; END_VAR
END_METHOD

METHOD M_SetParameter : BOOL
VAR_INPUT i_nAddress : WORD; i_wRawValue : WORD; END_VAR
END_METHOD

END_INTERFACE

// ---- 90_Project/PRG_Fast.TcPOU
PROGRAM PRG_Fast		// 빠른 계측 태스크에서 부름 (선택, 별도 코어 가능). 전력계를 빠르게 읽어야 하는 현장만
VAR
END_VAR

(* 자리만. 할 일
   - 빠른 계측 FB를 부르고 결과를 GVL_IF 계측 칸에 다 쓴 뒤 GVL_IF.g_nFastSeq를 1 올림
   - MAIN 쪽은 계측기 드라이버(I_Meter)가 GVL_IF에서 읽어 FB_Snapshot에 넘김
   - 계측 FB 인스턴스(I/O 연결 있음)는 이 PRG의 VAR에 선언 → I/O가 FastTask 주기로 갱신됨
     GVL에 두면 선언 위에 {attribute 'TcContextName' := 'FastTask'} 필요 (안 붙이면 PlcTask 주기로 갱신됨, 헬리오스 SETTING_VALUE 참고) *)
;

END_PROGRAM

// ---- 90_Project/PRG_Mqtt.TcPOU
PROGRAM PRG_Mqtt		// MqttTask에서 부름. 보고 올리기·명령 받기 (MQTT 담당자 영역)
(* - MAIN의 FB나 GVL_SITE·GVL_PERSIST를 직접 읽거나 쓰지 않는다 (GVL_SITE 상수 TEST_MODE·MQTT_SET만 읽음). 주고받기는 GVL_IF만
   - MQTT 클라이언트 FB 인스턴스(브로커 3개)는 FB_MqttMain 안에 있고 여기서만 부른다. 접속 설정은 GVL_SITE.MQTT_SET
   - 명령: 받은 command 레코드를 FB_EmsCommand(명령 핸들러)가 Std 명령으로 해석 → GVL_IF.g_stEmsCmd에 쓰고 번호(g_nCmdSeq)를 올림 → MAIN이 FB_SrcEms로 받음
   - 보고: 시험 모드면 먼저 더미 값(PRG_MqttTestData)을 채우고, MAIN이 GVL_IF.g_stReport에 채운 매핑된 PCS·BAT 레코드(A_Report)를 그 위에 덮어씀. 매핑이 없는 장치·토픽은 더미 그대로 *)
VAR
	nUpsConfigRxCount : UDINT; // last handed-over config/ups receive count
	fbMqttMain		: FB_MqttMain;		// 발행·구독 (브로커 3개)
	sInstance		: STRING(4);			// ClientId 꼬리표 (이중화일 때 역할로 정함)
	bRoleReady		: BOOL;				// 이중화 역할이 정해짐 (안 쓰면 항상 TRUE)
	fbEmsCommand	: FB_EmsCommand;		// 명령 핸들러
	fbGatePcs		: FB_EmsCmdGate;		// command/pcs 중복 거르기·Delay 대기 [2026-11-12]
	fbGateBat		: FB_EmsCmdGate;		// command/bat
	fbGateUps		: FB_EmsCmdGate;		// command/ups
	stRptCopy		: ST_IfReport;		// 보고 칸의 마지막 일관된 복사본
 stRptCandidate : ST_IfReport; // 복사 중인 보고값
	nRptSeq			: UDINT;
	bRptValid		: BOOL;
	nRxTotal		: UDINT;				// command 메시지 수신 누계 (브로커 3개 합)
	i				: UINT;
	(* [9-21 수정 2026-11-04: 추가] EMS config → GVL_IF, 실제 설정 echo ← GVL_IF *)
	stCfgOut		: ST_IfEmsCfg;		// GVL_IF.g_stEmsCfg에 올릴 칸 (마지막 레코드·번호 유지)
	nPrevPcsCfg		: UDINT;
	nPrevBatCfg		: UDINT;
	bCfgNew			: BOOL;
	k				: UDINT;
	nRec			: UDINT;
	nDev			: UINT;
	stPcsRec		: ST_PcsConfig_Rx;
	stBatRec		: ST_BatConfig_Rx;
	stCfgEchoCopy	: ST_IfEmsCfgEcho;
	nCfgEchoSeq		: UDINT;
END_VAR

(* 1. 발행 패킷 장치 번호, 시험 모드면 더미 발행 값 *)
PRG_PublishDeviceNo();
IF GVL_SITE.TEST_MODE THEN
	PRG_MqttTestData();
END_IF

(* 1-2. 보고: MAIN이 GVL_IF에 채운 PCS·BAT 레코드를 번호를 확인하며 복사해 발행 구조체에 넣음 (더미 위에 덮어씀).
   번호가 홀수 = 쓰는 중, 복사 전후 번호가 다름 = 복사 중에 바뀜 → 이번 스캔은 지난 복사본 그대로 *)
nRptSeq := GVL_IF.g_nReportSeq;
IF (nRptSeq AND 1) = 0 AND nRptSeq <> 0 THEN
	stRptCandidate := GVL_IF.g_stReport;
	IF GVL_IF.g_nReportSeq = nRptSeq THEN
  stRptCopy := stRptCandidate;
		bRptValid := TRUE;
	END_IF
END_IF
IF bRptValid THEN
	FOR i := 1 TO GVL_PARAM.PCS_COUNT DO
		IF stRptCopy.abPcsMapped[i] THEN
			g_stPcsPublish.Devices[i - 1] := stRptCopy.astPcs[i];
			g_stPcsPublish.Devices[i - 1].DeviceIndex := UINT_TO_UDINT(i);
		END_IF
	END_FOR
 FOR i := 1 TO GVL_PARAM.BMS_COUNT DO
  IF stRptCopy.abBatMapped[i] THEN
   g_stBatPublish.Devices[i - 1] := stRptCopy.astBat[i];
   g_stBatPublish.Devices[i - 1].DeviceIndex := UINT_TO_UDINT(i);
  END_IF
 END_FOR
 FOR i := 1 TO GVL_PARAM.RACK_COUNT DO
  IF stRptCopy.abBatMapped[(i - 1) / GVL_PARAM.RACKS_PER_BMS + 1] THEN
   g_stRackPublish.Devices[i - 1] := stRptCopy.astRack[i];
  END_IF
 END_FOR
 FOR i := 1 TO GVL_PARAM.BAT_MODULE_COUNT DO
  IF stRptCopy.abBatMapped[(i - 1) / (GVL_PARAM.RACKS_PER_BMS * GVL_PARAM.MODULES_PER_RACK) + 1] THEN
   g_stModulePublish.Devices[i - 1] := stRptCopy.astModule[i];
  END_IF
 END_FOR
 FOR i := 1 TO GVL_PARAM.UPS_COUNT DO
  IF stRptCopy.abUpsMapped[i] THEN
   g_stUpsPublish.Devices[i - 1] := stRptCopy.astUps[i];
   g_stUpsPublish.Devices[i - 1].DeviceIndex := UINT_TO_UDINT(i); // 번호 1부터
  END_IF
 END_FOR
 FOR i := 1 TO GVL_PARAM.IMD_COUNT DO
  IF stRptCopy.abImdMapped[i] THEN
   g_stImdPublish.Devices[i - 1] := stRptCopy.astImd[i];
   g_stImdPublish.Devices[i - 1].DeviceIndex := UINT_TO_UDINT(i); // 번호 1부터
  END_IF
 END_FOR
 FOR i := 1 TO GVL_PARAM.FIRE_COUNT DO
  IF stRptCopy.abFireMapped[i] THEN
   g_stFirePublish.Devices[i - 1] := stRptCopy.astFire[i]; // 번호 1부터 (MAIN이 채움)
  END_IF
 END_FOR
 FOR i := 1 TO GVL_PARAM.TEMP_COUNT DO
  IF stRptCopy.abTempMapped[i] THEN
   g_stTempPublish.Devices[i - 1] := stRptCopy.astTemp[i]; // 시험 더미 위에 덮어씀
  END_IF
 END_FOR
END_IF

(* 1-3. config echo: MAIN이 GVL_IF에 채운 실제 설정을 번호를 확인하며 복사 → GVL_MQTT applied 칸 (FB_MqttMain이 config echo로 발행) [9-21 수정 2026-11-04: 추가] *)
nCfgEchoSeq := GVL_IF.g_nCfgEchoSeq;
IF (nCfgEchoSeq AND 1) = 0 AND nCfgEchoSeq <> 0 THEN
	stCfgEchoCopy := GVL_IF.g_stEmsCfgEcho;
	IF GVL_IF.g_nCfgEchoSeq = nCfgEchoSeq THEN
		GVL_MQTT.g_astPcsConfigApplied	:= stCfgEchoCopy.astPcs;
		GVL_MQTT.g_astBatConfigApplied	:= stCfgEchoCopy.astBat;
		GVL_MQTT.g_bConfigApplied		:= TRUE;
	END_IF
END_IF

(* 2. 발행·구독 (브로커 3개) *)
// 이중화: 두 PLC가 같은 사이트·같은 ClientId로 접속하면 브로커가 서로 끊으므로 역할로 ClientId를 구분. 발행은 Active만, 구독은 두 PLC 모두
IF GVL_SITE.RED_SET.bUse THEN
	CASE GVL_IF.g_eRedRole OF
	E_RedRole.Primary:		sInstance := '-P'; bRoleReady := TRUE;
	E_RedRole.Secondary:	sInstance := '-S'; bRoleReady := TRUE;
	ELSE					sInstance := '';   bRoleReady := FALSE;	// 읽는 중·설정 오류: 접속하지 않음
	END_CASE
ELSE
	sInstance	:= '';
	bRoleReady	:= TRUE;
END_IF
fbMqttMain(	i_stSet		:= GVL_SITE.MQTT_SET,
			i_sInstance	:= sInstance,
			i_bPublish	:= GVL_IF.g_bRedActive,
			i_bReady	:= bRoleReady);
GVL_IF.g_abBrokerUse	:= fbMqttMain.q_abBrokerUse;	// [9번 수정 2026-11-09: 추가] 브로커 접속 상태 → MAIN (FB_BrokerWatch)
GVL_IF.g_abBrokerConn	:= fbMqttMain.q_abBrokerConn;

// config/ups is raw receipt staging only. No setting application or hardware request.
IF GVL_MQTT.g_anCfgRxCount[4]<>nUpsConfigRxCount THEN
 nUpsConfigRxCount:=GVL_MQTT.g_anCfgRxCount[4];
 GVL_IF.g_nUpsConfigSeq:=GVL_IF.g_nUpsConfigSeq+1;
 GVL_IF.g_stUpsConfigRx.astConfig:=GVL_MQTT.g_astUpsConfig;
 GVL_IF.g_stUpsConfigRx.nRxCount:=nUpsConfigRxCount;
 GVL_IF.g_nUpsConfigSeq:=GVL_IF.g_nUpsConfigSeq+1;
END_IF

(* 2-1. 로거 발행 시험 (시험 모드. 버튼을 누를 때만 로그를 남김, 결과는 PRG_TestLogger 머리말) *)
IF GVL_SITE.TEST_MODE THEN
	PRG_TestLogger();
END_IF

(* 3. 수신 시험 기록 (시험 모드. 명령 핸들러가 CommandType을 지우기 전의 사본) *)
IF GVL_SITE.TEST_MODE THEN
	PRG_MqttTestData.A_HandleRx();
END_IF

(* 3-1. 명령 앞단 (인터페이스 100.Command 2026-11-12): 같은 SequenceNumber 버리기, Delay(ms)만큼 기다렸다가 핸들러에 넘김 *)
fbGatePcs(iq_astRec := g_astPcsCommand);
fbGateBat(iq_astRec := g_astBatCommand);
fbGateUps(iq_astRec := g_astUpsCommand);

(* 4. 명령 핸들러: command 레코드 → Std 명령. 바뀌었으면 GVL_IF에 올림 (쓰기 전 번호 홀수, 끝나면 짝수) *)
nRxTotal := 0;
FOR i := 1 TO GVL_MQTT.COMMAND_TOPIC_COUNT DO
	nRxTotal := nRxTotal + g_anCmdRxCount[i];
END_FOR
fbEmsCommand(	i_nRxCount			:= nRxTotal,
				iq_astPcsCommand	:= g_astPcsCommand,
				iq_astBatCommand	:= g_astBatCommand);
IF fbEmsCommand.q_bChanged THEN
	GVL_IF.g_nCmdSeq := GVL_IF.g_nCmdSeq + 1;
	GVL_IF.g_stEmsCmd := fbEmsCommand.q_stCmd;
	GVL_IF.g_nCmdSeq := GVL_IF.g_nCmdSeq + 1;
END_IF

(* 5. EMS config(pcs·bat) → GVL_IF.g_stEmsCfg [9-21 수정 2026-11-04: 추가]. 새 메시지(수신 횟수가 바뀜)의 레코드를 칸(DeviceId, 1부터 [1부터 2026-11-10])에 넣고 그 칸 번호를 올림.
   실제로 받은 레코드(GVL_MQTT.g_anCfgRxRecords)까지만 봄. 반영은 MAIN (FB_EmsConfigApply)
   [21번 수정 2026-11-09: is_available이 모두 0인 레코드도 넘김 (기본값으로 반영 = 한도 해제). 원래는 그런 레코드를 빈 칸으로 보고 건너뜀
    → 빈 칸은 받은 레코드 수로 거름 (헤더 DeviceCount가 실제보다 크면 그 뒤 칸은 0으로 채워져 PCS 1로 보이므로)] *)
bCfgNew := FALSE;
IF GVL_MQTT.g_anCfgRxCount[1] <> nPrevPcsCfg THEN
	nPrevPcsCfg := GVL_MQTT.g_anCfgRxCount[1];
	nRec := MIN(MIN(GVL_MQTT.g_stPcsConfigWireIn.Header.DeviceCount, GVL_MQTT.g_anCfgRxRecords[1]), UINT_TO_UDINT(GVL_PARAM.PCS_COUNT));
	FOR k := 1 TO nRec DO
		stPcsRec := GVL_MQTT.g_stPcsConfigWireIn.Records[k - 1];
		IF stPcsRec.DeviceId >= 1 AND stPcsRec.DeviceId <= UINT_TO_UDINT(GVL_PARAM.PCS_COUNT) THEN
			nDev := UDINT_TO_UINT(stPcsRec.DeviceId);
			stCfgOut.astPcs[nDev]	:= stPcsRec;
			stCfgOut.anPcsSeq[nDev]	:= stCfgOut.anPcsSeq[nDev] + 1;
			bCfgNew := TRUE;
		END_IF
	END_FOR
END_IF
IF GVL_MQTT.g_anCfgRxCount[2] <> nPrevBatCfg THEN
	nPrevBatCfg := GVL_MQTT.g_anCfgRxCount[2];
	nRec := MIN(MIN(GVL_MQTT.g_stBatConfigWireIn.Header.DeviceCount, GVL_MQTT.g_anCfgRxRecords[2]), UINT_TO_UDINT(GVL_PARAM.BMS_COUNT));
	FOR k := 1 TO nRec DO
		stBatRec := GVL_MQTT.g_stBatConfigWireIn.Records[k - 1];
		IF stBatRec.DeviceId >= 1 AND stBatRec.DeviceId <= UINT_TO_UDINT(GVL_PARAM.BMS_COUNT) THEN
			nDev := UDINT_TO_UINT(stBatRec.DeviceId);
			stCfgOut.astBat[nDev]	:= stBatRec;
			stCfgOut.anBatSeq[nDev]	:= stCfgOut.anBatSeq[nDev] + 1;
			bCfgNew := TRUE;
		END_IF
	END_FOR
END_IF
IF bCfgNew THEN
	GVL_IF.g_nCfgSeq := GVL_IF.g_nCfgSeq + 1;
	GVL_IF.g_stEmsCfg := stCfgOut;
	GVL_IF.g_nCfgSeq := GVL_IF.g_nCfgSeq + 1;
END_IF

(* 6. UPS 명령 (명세 WR-UPS-01): command/ups 레코드 → GVL_IF.g_astUpsCmd. 받은 레코드는 지움. MAIN.fbUpsCommand가 실행 *)
FOR i := 0 TO GVL_PARAM.UPS_COUNT - 1 DO
	IF g_astUpsCommand[i].CommandType <> 0 THEN
		GVL_IF.g_nUpsCmdSeq := GVL_IF.g_nUpsCmdSeq + 1;	// 홀수 = 쓰는 중
		GVL_IF.g_astUpsCmd[i + 1].nType := g_astUpsCommand[i].CommandType;
		GVL_IF.g_astUpsCmd[i + 1].nSeq := GVL_IF.g_astUpsCmd[i + 1].nSeq + 1;
		GVL_IF.g_nUpsCmdSeq := GVL_IF.g_nUpsCmdSeq + 1;	// 짝수 = 끝
		g_astUpsCommand[i].CommandType := 0;
	END_IF
END_FOR

END_PROGRAM

// ---- 20_Module/Mqtt/FB_MqttMain.TcPOU
FUNCTION_BLOCK FB_MqttMain		// MQTT 보고·명령 로직: 시각 문자열, 발행·구독 토픽 표, 브로커 3개(Cloud·Local·Azure) 발행·구독, 로거 이벤트 발행 (PRG_Mqtt가 부름. 접속 설정은 i_stSet = GVL_SITE.MQTT_SET)
VAR_INPUT
	i_stSet				: ST_MqttSet;		// 접속 설정 (사이트 번호·브로커·계정)
	i_sInstance			: STRING(4) := '';	// ClientId 뒤에 붙임. 이중화: Primary '-P', Secondary '-S' (두 PLC가 같은 ClientId면 브로커가 서로 끊음)
	i_bPublish			: BOOL := TRUE;		// 발행 허가 (이중화: Active만 발행. 구독은 두 PLC 모두)
	i_bReady			: BOOL := TRUE;		// 접속 시작 허가 (이중화: 역할이 정해진 뒤)
END_VAR
VAR_OUTPUT
	q_abBrokerUse		: ARRAY[1..3] OF BOOL;	// 쓰는 브로커 (1 Cloud, 2 Local, 3 Azure = i_stSet bUse) [9번 수정 2026-11-09: 추가]
	q_abBrokerConn		: ARRAY[1..3] OF BOOL;	// 구독 클라이언트가 접속됨 (쓰지 않는 브로커·접속 시작 전은 FALSE)
END_VAR
VAR
	(* ---------- 토픽 표 ---------- *)
	bTableInit			: BOOL;
	astPubDeviceTable	: ARRAY[1..GVL_MQTT.DEVICE_TOPIC_COUNT] OF ST_MqttPubEntry;
	astPubConfigTable	: ARRAY[1..GVL_MQTT.CONFIG_TOPIC_COUNT] OF ST_MqttPubEntry;
	astSubCommandTable	: ARRAY[1..GVL_MQTT.COMMAND_TOPIC_COUNT] OF ST_MqttSubEntry;
	astSubConfigTable	: ARRAY[1..GVL_MQTT.CONFIG_TOPIC_COUNT] OF ST_MqttSubEntry;

	(* 토픽별 수신 버퍼: 헤더 + 그 토픽의 최대 레코드 수 (config pcs·bat은 GVL_MQTT 수신 패킷을 버퍼로 씀) *)
	anRxPcsCommand		: ARRAY[0..(SIZEOF(ST_MqttCommandHeader) + SIZEOF(ST_MqttCommand_Rx) * GVL_PARAM.PCS_COUNT - 1)] OF BYTE;
	anRxBatCommand		: ARRAY[0..(SIZEOF(ST_MqttCommandHeader) + SIZEOF(ST_MqttCommand_Rx) * GVL_PARAM.BMS_COUNT - 1)] OF BYTE;
	anRxUpsCommand		: ARRAY[0..(SIZEOF(ST_MqttCommandHeader) + SIZEOF(ST_MqttCommand_Rx) * GVL_PARAM.UPS_COUNT - 1)] OF BYTE;
	anRxProtectionConfig : ARRAY[0..(SIZEOF(ST_MqttCommandHeader) + SIZEOF(ST_ProtectionConfig_Rx) - 1)] OF BYTE;

	(* ---------- 브로커 ---------- *)
	fbCloudSub			: FB_MqttSubscribe;
	fbCloudPub			: FB_MqttPublish;
	fbLocalSub			: FB_MqttSubscribe;
	fbLocalPub			: FB_MqttPublish;
	fbAzureSub			: FB_MqttSubscribe;
	fbAzurePub			: FB_MqttPublish;
	tonStartDelay		: TON := (PT := T#10S);		// 기동 뒤 통신 시작 지연

	(* ---------- 시각 ---------- *)
	fbLocalTime			: FB_LocalSystemTime := (sNetID := '', bEnable := TRUE);
	sTimeStamp			: STRING(23);		// '2024-09-04 11:11:11.123' (보고 헤더·DB 저장 시각)

	(* ---------- 수신 합산 (브로커 3개 → GVL_MQTT) ---------- *)
	i					: UINT;
	anPrevCmdCount		: ARRAY[1..3, 1..GVL_MQTT.COMMAND_TOPIC_COUNT] OF UDINT;	// 1 Cloud, 2 Local, 3 Azure
	anPrevCfgCount		: ARRAY[1..3, 1..GVL_MQTT.CONFIG_TOPIC_COUNT] OF UDINT;

	(* ---------- 로거 (이벤트 로그 → pms_log 토픽, 20_Module/Mqtt/Logger) ---------- *)
	fbLogger			: FB_MqttLoggerListener;
	anLoggerNext		: ARRAY[1..3] OF UDINT := [1, 1, 1];	// 브로커별 다음에 보낼 이벤트 번호 (1 Cloud, 2 Local, 3 Azure)
	stLoggerPacket		: ST_LoggerPublish_V1;
	nUtcOffset			: LINT;		// 현지 시각 − UTC (100 ns). 로거 시각(UTC)을 현지 시각으로 바꿀 때 씀
	bUtcOffsetValid		: BOOL;
	stLocalFileTime		: T_FILETIME;
	nLocalFileTime		: ULINT;
	nOffsetRaw			: LINT;
END_VAR
VAR CONSTANT
	OFFSET_STEP			: LINT := 9000000000;	// 시간대 단위 15분 (100 ns). 두 시각을 읽는 사이의 차이를 반올림으로 없앰
END_VAR

(* 1. 시각 문자열 *)
fbLocalTime();
A_MakeTimeStamp();

(* 2. 토픽 표 (처음 한 번) *)
IF NOT bTableInit THEN
	A_InitPublishTable();
	A_InitSubscribeTable();
	bTableInit := TRUE;
END_IF
A_MapPublishHeader();

(* 2-1. 로거 이벤트 받기: 접속 지연과 상관없이 처음부터 (기동 직후 로그도 큐에 쌓였다가 접속하면 나감) *)
fbLogger.M_Cycle(i_nUtcOffset := nUtcOffset, i_bTimeValid := bUtcOffsetValid);

(* 3. 브로커 발행·구독 *)
tonStartDelay(IN := TRUE);
IF tonStartDelay.Q AND i_bReady THEN
	IF i_stSet.stCloud.bUse THEN
		fbCloudPub(i_sConnLabel := 'Cloud', i_nSiteId := i_stSet.nSiteId, i_sHost := i_stSet.stCloud.sHost, i_nPort := i_stSet.stCloud.nPort, i_sUserName := i_stSet.sUserName, i_sUserPassword := i_stSet.sUserPassword, i_astDeviceTable := astPubDeviceTable, i_sInstance := i_sInstance, i_bPublish := i_bPublish, i_astConfigTable := astPubConfigTable);
		fbCloudSub(i_nSiteId := i_stSet.nSiteId, i_sHost := i_stSet.stCloud.sHost, i_nPort := i_stSet.stCloud.nPort, i_sUserName := i_stSet.sUserName, i_sUserPassword := i_stSet.sUserPassword, i_astCommandTable := astSubCommandTable, i_sInstance := i_sInstance, i_astConfigTable := astSubConfigTable);
	END_IF
	IF i_stSet.stLocal.bUse THEN
		fbLocalPub(i_sConnLabel := 'local', i_nSiteId := i_stSet.nSiteId, i_sHost := i_stSet.stLocal.sHost, i_nPort := i_stSet.stLocal.nPort, i_sUserName := i_stSet.sUserName, i_sUserPassword := i_stSet.sUserPassword, i_astDeviceTable := astPubDeviceTable, i_sInstance := i_sInstance, i_bPublish := i_bPublish, i_astConfigTable := astPubConfigTable);
		fbLocalSub(i_nSiteId := i_stSet.nSiteId, i_sHost := i_stSet.stLocal.sHost, i_nPort := i_stSet.stLocal.nPort, i_sUserName := i_stSet.sUserName, i_sUserPassword := i_stSet.sUserPassword, i_astCommandTable := astSubCommandTable, i_sInstance := i_sInstance, i_astConfigTable := astSubConfigTable);
	END_IF
	IF i_stSet.stAzure.bUse THEN
		fbAzurePub(i_sConnLabel := 'Azure', i_nSiteId := i_stSet.nSiteId, i_sHost := i_stSet.stAzure.sHost, i_nPort := i_stSet.stAzure.nPort, i_sUserName := i_stSet.sUserName, i_sUserPassword := i_stSet.sUserPassword, i_astDeviceTable := astPubDeviceTable, i_sInstance := i_sInstance, i_bPublish := i_bPublish, i_astConfigTable := astPubConfigTable);
		fbAzureSub(i_nSiteId := i_stSet.nSiteId, i_sHost := i_stSet.stAzure.sHost, i_nPort := i_stSet.stAzure.nPort, i_sUserName := i_stSet.sUserName, i_sUserPassword := i_stSet.sUserPassword, i_astCommandTable := astSubCommandTable, i_sInstance := i_sInstance, i_astConfigTable := astSubConfigTable);
	END_IF

	A_MergeRxCount();
	A_PublishLogger();
END_IF
// [9번 수정 2026-11-09: 추가] 브로커 접속 상태 (PRG_Mqtt → GVL_IF → MAIN FB_BrokerWatch)
q_abBrokerUse[1]	:= i_stSet.stCloud.bUse;
q_abBrokerUse[2]	:= i_stSet.stLocal.bUse;
q_abBrokerUse[3]	:= i_stSet.stAzure.bUse;
q_abBrokerConn[1]	:= i_stSet.stCloud.bUse AND tonStartDelay.Q AND i_bReady AND fbCloudSub.q_bConnected;
q_abBrokerConn[2]	:= i_stSet.stLocal.bUse AND tonStartDelay.Q AND i_bReady AND fbLocalSub.q_bConnected;
q_abBrokerConn[3]	:= i_stSet.stAzure.bUse AND tonStartDelay.Q AND i_bReady AND fbAzureSub.q_bConnected;

ACTION A_InitPublishTable:
astPubDeviceTable[1].sTopic          := 'pms';
astPubDeviceTable[1].pDeviceSrc       := ADR(g_stPmsPublish.Devices);
astPubDeviceTable[1].nDeviceElemSize  := SIZEOF(ST_PmsPublish_V1);
astPubDeviceTable[1].nDeviceCount     := 1;
astPubDeviceTable[1].pStaging         := ADR(g_stPmsPublish);
astPubDeviceTable[1].nStagingSize     := SIZEOF(g_stPmsPublish);
astPubDeviceTable[1].sCategory       := '';

astPubDeviceTable[2].sTopic          := 'pcs';
astPubDeviceTable[2].pDeviceSrc       := ADR(g_stPcsPublish.Devices);
astPubDeviceTable[2].nDeviceElemSize  := SIZEOF(ST_PcsPublish_V1);
astPubDeviceTable[2].nDeviceCount     := UINT_TO_UDINT(GVL_PARAM.INSTALLED_PCS_COUNT);
astPubDeviceTable[2].pStaging         := ADR(g_stPcsPublish);
astPubDeviceTable[2].nStagingSize     := SIZEOF(g_stPcsPublish);
astPubDeviceTable[2].sCategory       := '';

astPubDeviceTable[3].sTopic          := 'bat';
astPubDeviceTable[3].pDeviceSrc       := ADR(g_stBatPublish.Devices);
astPubDeviceTable[3].nDeviceElemSize  := SIZEOF(ST_BatPublish_V1);
astPubDeviceTable[3].nDeviceCount     := UINT_TO_UDINT(GVL_PARAM.BMS_COUNT);
astPubDeviceTable[3].pStaging         := ADR(g_stBatPublish);
astPubDeviceTable[3].nStagingSize     := SIZEOF(g_stBatPublish);
astPubDeviceTable[3].sCategory       := '';


astPubDeviceTable[4].sTopic          := 'rack';
astPubDeviceTable[4].pDeviceSrc       := ADR(g_stRackPublish.Devices);
astPubDeviceTable[4].nDeviceElemSize  := SIZEOF(ST_RackPublish_V1);
astPubDeviceTable[4].nDeviceCount     := UINT_TO_UDINT(GVL_PARAM.RACK_COUNT);
astPubDeviceTable[4].pStaging         := ADR(g_stRackPublish);
astPubDeviceTable[4].nStagingSize     := SIZEOF(g_stRackPublish);
astPubDeviceTable[4].sCategory       := '';

astPubDeviceTable[5].sTopic          := 'pv_meter';
astPubDeviceTable[5].pDeviceSrc       := ADR(g_stPvPublish.Devices);
astPubDeviceTable[5].nDeviceElemSize  := SIZEOF(ST_PvPublish_V1);
astPubDeviceTable[5].nDeviceCount     := UINT_TO_UDINT(GVL_PARAM.PV_COUNT);
astPubDeviceTable[5].pStaging         := ADR(g_stPvPublish);
astPubDeviceTable[5].nStagingSize     := SIZEOF(g_stPvPublish);
astPubDeviceTable[5].sCategory       := '';

astPubDeviceTable[6].sTopic          := 'ess_meter';
astPubDeviceTable[6].pDeviceSrc       := ADR(g_stEssPublish.Devices);
astPubDeviceTable[6].nDeviceElemSize  := SIZEOF(ST_EssPublish_V1);
astPubDeviceTable[6].nDeviceCount     := UINT_TO_UDINT(GVL_PARAM.ESS_COUNT);
astPubDeviceTable[6].pStaging         := ADR(g_stEssPublish);
astPubDeviceTable[6].nStagingSize     := SIZEOF(g_stEssPublish);
astPubDeviceTable[6].sCategory       := '';

astPubDeviceTable[7].sTopic          := 'temperature_sensor';
astPubDeviceTable[7].pDeviceSrc       := ADR(g_stTempPublish.Devices);
astPubDeviceTable[7].nDeviceElemSize  := SIZEOF(ST_TempPublish_V1);
astPubDeviceTable[7].nDeviceCount     := UINT_TO_UDINT(GVL_PARAM.TEMP_COUNT);
astPubDeviceTable[7].pStaging         := ADR(g_stTempPublish);
astPubDeviceTable[7].nStagingSize     := SIZEOF(g_stTempPublish);
astPubDeviceTable[7].sCategory       := '';

astPubDeviceTable[8].sTopic          := 'airconditioner'; //공조기
astPubDeviceTable[8].pDeviceSrc       := ADR(g_stAirConditionerPublish.Devices);
astPubDeviceTable[8].nDeviceElemSize  := SIZEOF(ST_AirConditionerPublish_V1);
astPubDeviceTable[8].nDeviceCount     := UINT_TO_UDINT(GVL_PARAM.AIR_CONDITIONER_COUNT);
astPubDeviceTable[8].pStaging         := ADR(g_stAirConditionerPublish);
astPubDeviceTable[8].nStagingSize     := SIZEOF(g_stAirConditionerPublish);
astPubDeviceTable[8].sCategory       := '';

astPubDeviceTable[9].sTopic := 'ups';
astPubDeviceTable[9].sCategory := '';
astPubDeviceTable[9].pDeviceSrc := ADR(g_stUpsPublish.Devices);
astPubDeviceTable[9].nDeviceElemSize := SIZEOF(ST_UpsPublish_V1);
astPubDeviceTable[9].nDeviceCount := SEL(GVL_MQTT.UPS_REPORT_ENABLED,UDINT#0,UINT_TO_UDINT(GVL_PARAM.UPS_COUNT));
astPubDeviceTable[9].pStaging := ADR(g_stUpsPublish);
astPubDeviceTable[9].nStagingSize := SIZEOF(g_stUpsPublish);
astPubDeviceTable[10].sTopic := 'module';
astPubDeviceTable[10].sCategory := '';
astPubDeviceTable[10].pDeviceSrc := ADR(g_stModulePublish.Devices);
astPubDeviceTable[10].nDeviceElemSize := SIZEOF(ST_ModulePublish_V1);
astPubDeviceTable[10].nDeviceCount := SEL(GVL_MQTT.MODULE_REPORT_ENABLED,UDINT#0,UINT_TO_UDINT(GVL_PARAM.BAT_MODULE_COUNT));
astPubDeviceTable[10].pStaging := ADR(g_stModulePublish);
astPubDeviceTable[10].nStagingSize := SIZEOF(g_stModulePublish);
astPubDeviceTable[11].sTopic := 'imd'; // IMD 절연감시
astPubDeviceTable[11].sCategory := '';
astPubDeviceTable[11].pDeviceSrc := ADR(g_stImdPublish.Devices);
astPubDeviceTable[11].nDeviceElemSize := SIZEOF(ST_ImdPublish_V1);
astPubDeviceTable[11].nDeviceCount := SEL(GVL_MQTT.IMD_REPORT_ENABLED,UDINT#0,UINT_TO_UDINT(GVL_PARAM.IMD_COUNT));
astPubDeviceTable[11].pStaging := ADR(g_stImdPublish);
astPubDeviceTable[11].nStagingSize := SIZEOF(g_stImdPublish);
astPubDeviceTable[12].sTopic := 'fire_detector'; // 화재감지기 (OffGas 양식, 이름 잠정)
astPubDeviceTable[12].sCategory := '';
astPubDeviceTable[12].pDeviceSrc := ADR(g_stFirePublish.Devices);
astPubDeviceTable[12].nDeviceElemSize := SIZEOF(ST_FirePublish_V1);
astPubDeviceTable[12].nDeviceCount := SEL(GVL_MQTT.FIRE_REPORT_ENABLED,UDINT#0,UINT_TO_UDINT(GVL_PARAM.FIRE_COUNT));
astPubDeviceTable[12].pStaging := ADR(g_stFirePublish);
astPubDeviceTable[12].nStagingSize := SIZEOF(g_stFirePublish);
astPubConfigTable[4].sCategory := 'config';
astPubConfigTable[4].sTopic := 'ups';
astPubConfigTable[4].pDeviceSrc := ADR(g_stUpsConfigEcho.Records);
astPubConfigTable[4].nDeviceElemSize := SIZEOF(ST_UpsConfig_Rx);
astPubConfigTable[4].nDeviceCount := UINT_TO_UDINT(GVL_PARAM.UPS_COUNT);
astPubConfigTable[4].pStaging := ADR(g_stUpsConfigEcho);
astPubConfigTable[4].nStagingSize := SIZEOF(g_stUpsConfigEcho);

(* config echo *)
astPubConfigTable[1].sCategory       := 'config';
astPubConfigTable[1].sTopic          := 'pcs';
astPubConfigTable[1].pDeviceSrc      := ADR(g_stPcsConfigEcho.Records);
astPubConfigTable[1].nDeviceElemSize := SIZEOF(ST_PcsConfig_Rx);
astPubConfigTable[1].nDeviceCount    := UINT_TO_UDINT(GVL_PARAM.INSTALLED_PCS_COUNT);
astPubConfigTable[1].pStaging        := ADR(g_stPcsConfigEcho);
astPubConfigTable[1].nStagingSize    := SIZEOF(g_stPcsConfigEcho);

astPubConfigTable[2].sCategory       := 'config';
astPubConfigTable[2].sTopic          := 'bat';
astPubConfigTable[2].pDeviceSrc      := ADR(g_stBatConfigEcho.Records);
astPubConfigTable[2].nDeviceElemSize := SIZEOF(ST_BatConfig_Rx);
astPubConfigTable[2].nDeviceCount    := UINT_TO_UDINT(GVL_PARAM.BMS_COUNT);
astPubConfigTable[2].pStaging        := ADR(g_stBatConfigEcho);
astPubConfigTable[2].nStagingSize    := SIZEOF(g_stBatConfigEcho);

astPubConfigTable[3].sCategory       := 'config';
astPubConfigTable[3].sTopic          := 'protection';
astPubConfigTable[3].pDeviceSrc      := ADR(g_stProtectionConfigEcho.Record);	// [결함 12 수정 2026-11-04: 원래 g_stProtectionConfigWireIn]
astPubConfigTable[3].nDeviceElemSize := SIZEOF(ST_ProtectionConfig_Rx);
astPubConfigTable[3].nDeviceCount    := 1;
astPubConfigTable[3].pStaging        := ADR(g_stProtectionConfigEcho);
astPubConfigTable[3].nStagingSize    := SIZEOF(g_stProtectionConfigEcho);
END_ACTION

ACTION A_InitSubscribeTable:
(*command*)
astSubCommandTable[1].sCategory   := 'command';
astSubCommandTable[1].sTopic      := 'pcs';
astSubCommandTable[1].bIndexed    := TRUE;
astSubCommandTable[1].pDestArray  := ADR(g_astPcsCommand);
astSubCommandTable[1].nElementSize:= SIZEOF(ST_MqttCommand_Rx);
astSubCommandTable[1].nDeviceCapacity    := UINT_TO_UDINT(GVL_PARAM.PCS_COUNT);
astSubCommandTable[1].pRxBuffer      := ADR(anRxPcsCommand);
astSubCommandTable[1].nRxBufferSize  := SIZEOF(anRxPcsCommand);
astSubCommandTable[1].nMaxRecords     := (SIZEOF(anRxPcsCommand) - SIZEOF(ST_MqttCommandHeader)) / SIZEOF(ST_MqttCommand_Rx);
astSubCommandTable[1].nIndexOffset    := 4;	// SequenceNumber 뒤 DeviceIndex [2026-11-12]

astSubCommandTable[2].sCategory   := 'command';
astSubCommandTable[2].sTopic      := 'bat';
astSubCommandTable[2].bIndexed    := TRUE;
astSubCommandTable[2].pDestArray  := ADR(g_astBatCommand);
astSubCommandTable[2].nElementSize:= SIZEOF(ST_MqttCommand_Rx);
astSubCommandTable[2].nDeviceCapacity    := UINT_TO_UDINT(GVL_PARAM.BMS_COUNT);
astSubCommandTable[2].pRxBuffer      := ADR(anRxBatCommand);
astSubCommandTable[2].nRxBufferSize  := SIZEOF(anRxBatCommand);
astSubCommandTable[2].nMaxRecords     := (SIZEOF(anRxBatCommand) - SIZEOF(ST_MqttCommandHeader)) / SIZEOF(ST_MqttCommand_Rx);
astSubCommandTable[2].nIndexOffset    := 4;

astSubCommandTable[3].sCategory   := 'command';
astSubCommandTable[3].sTopic      := 'ups';
astSubCommandTable[3].bIndexed    := TRUE;
astSubCommandTable[3].pDestArray  := ADR(g_astUpsCommand);
astSubCommandTable[3].nElementSize:= SIZEOF(ST_MqttCommand_Rx);
astSubCommandTable[3].nDeviceCapacity    := UINT_TO_UDINT(GVL_PARAM.UPS_COUNT);
astSubCommandTable[3].pRxBuffer      := ADR(anRxUpsCommand);
astSubCommandTable[3].nRxBufferSize  := SIZEOF(anRxUpsCommand);
astSubCommandTable[3].nMaxRecords     := (SIZEOF(anRxUpsCommand) - SIZEOF(ST_MqttCommandHeader)) / SIZEOF(ST_MqttCommand_Rx);
astSubCommandTable[3].nIndexOffset    := 4;
// UPS 번호도 1부터: F_MqttDistribute.DEVICE_ID_BASE가 모든 토픽에 적용 (원래 여기서 nDeviceIdBase := 1) [1부터 2026-11-10]

astSubConfigTable[4].sCategory := 'config';
astSubConfigTable[4].sTopic := 'ups';
astSubConfigTable[4].bIndexed := TRUE;
astSubConfigTable[4].pDestArray := ADR(g_astUpsConfig);
astSubConfigTable[4].nElementSize := SIZEOF(ST_UpsConfig_Rx);
astSubConfigTable[4].nDeviceCapacity := UINT_TO_UDINT(GVL_PARAM.UPS_COUNT);
astSubConfigTable[4].pRxBuffer := ADR(g_stUpsConfigWireIn);
astSubConfigTable[4].nRxBufferSize := SIZEOF(g_stUpsConfigWireIn);
astSubConfigTable[4].nMaxRecords := UINT_TO_UDINT(GVL_PARAM.UPS_COUNT);
// UPS DeviceId 1부터: DEVICE_ID_BASE 적용 (원래 nDeviceIdBase := 1) [1부터 2026-11-10]

(*config*)
astSubConfigTable[1].sCategory   := 'config';
astSubConfigTable[1].sTopic      := 'pcs';
astSubConfigTable[1].bIndexed    := TRUE;
astSubConfigTable[1].pDestArray  := ADR(g_astPcsConfig);
astSubConfigTable[1].nElementSize:= SIZEOF(ST_PcsConfig_Rx);
astSubConfigTable[1].nDeviceCapacity    := UINT_TO_UDINT(GVL_PARAM.PCS_COUNT);
astSubConfigTable[1].pRxBuffer      := ADR(g_stPcsConfigWireIn);
astSubConfigTable[1].nRxBufferSize  := SIZEOF(g_stPcsConfigWireIn);
astSubConfigTable[1].nMaxRecords		:=(SIZEOF(g_stPcsConfigWireIn) - SIZEOF(ST_MqttCommandHeader)) / SIZEOF(ST_PcsConfig_Rx);

astSubConfigTable[2].sCategory   := 'config';
astSubConfigTable[2].sTopic      := 'bat';
astSubConfigTable[2].bIndexed    := TRUE;
astSubConfigTable[2].pDestArray  := ADR(g_astBatConfig);
astSubConfigTable[2].nElementSize:= SIZEOF(ST_BatConfig_Rx);
astSubConfigTable[2].nDeviceCapacity    := UINT_TO_UDINT(GVL_PARAM.BMS_COUNT);
astSubConfigTable[2].pRxBuffer      := ADR(g_stBatConfigWireIn);
astSubConfigTable[2].nRxBufferSize  := SIZEOF(g_stBatConfigWireIn);
astSubConfigTable[2].nMaxRecords		:=(SIZEOF(g_stBatConfigWireIn) - SIZEOF(ST_MqttCommandHeader)) / SIZEOF(ST_BatConfig_Rx);

astSubConfigTable[3].sCategory   := 'config';
astSubConfigTable[3].sTopic      := 'protection';
astSubConfigTable[3].bIndexed    := FALSE;		// DeviceIndex 없는 단일 레코드
astSubConfigTable[3].pDestArray  := ADR(g_stProtectionConfig);
astSubConfigTable[3].nElementSize:= SIZEOF(ST_ProtectionConfig_Rx);
astSubConfigTable[3].nDeviceCapacity    := 1;
astSubConfigTable[3].pRxBuffer      := ADR(g_stProtectionConfigWireIn);	// [결함 12 수정 2026-11-04: pcs·bat처럼 수신 버퍼 = WireIn (헤더 Location·UserName을 echo에 씀). 원래 ADR(anRxProtectionConfig)]
astSubConfigTable[3].nRxBufferSize  := SIZEOF(g_stProtectionConfigWireIn);	// [결함 12 수정 2026-11-04: 원래 SIZEOF(anRxProtectionConfig)]
astSubConfigTable[3].nMaxRecords     := (SIZEOF(g_stProtectionConfigWireIn) - SIZEOF(ST_MqttCommandHeader)) / SIZEOF(ST_ProtectionConfig_Rx);	// [결함 12 수정 2026-11-04: 원래 SIZEOF(anRxProtectionConfig)] // 결과적으로 1
END_ACTION

ACTION A_MakeTimeStamp:
(* 현지 시각 → '2024-09-04 11:11:11.123' (F_MqttTimeText).
   같이 현지 − UTC 차이를 구해 둔다 (로거 시각을 현지 시각으로 바꿀 때). 시간대는 15분 단위라 반올림.
   현지 시각을 아직 못 얻었으면(bValid FALSE) 지난 값 유지 *)
IF fbLocalTime.bValid THEN
	sTimeStamp := F_MqttTimeText(fbLocalTime.systemTime);

	stLocalFileTime := SYSTEMTIME_TO_FILETIME(fbLocalTime.systemTime);
	MEMCPY(destAddr := ADR(nLocalFileTime), srcAddr := ADR(stLocalFileTime), n := SIZEOF(nLocalFileTime));
	nOffsetRaw := ULINT_TO_LINT(nLocalFileTime) - ULINT_TO_LINT(F_GetSystemTime());
	IF nOffsetRaw >= 0 THEN
		nUtcOffset := ((nOffsetRaw + OFFSET_STEP / 2) / OFFSET_STEP) * OFFSET_STEP;
	ELSE
		nUtcOffset := -((((-nOffsetRaw) + OFFSET_STEP / 2) / OFFSET_STEP) * OFFSET_STEP);
	END_IF
	bUtcOffsetValid := TRUE;
END_IF
END_ACTION

ACTION A_MapPublishHeader:
g_stPmsPublish.Header.HeaderVersion := GVL_MQTT.HEADER_VERSION;
g_stPmsPublish.Header.DeviceVersion := GVL_MQTT.DEVICE_VERSION;
g_stPmsPublish.Header.SiteId        := i_stSet.nSiteId;
g_stPmsPublish.Header.DeviceCount   := 1;
g_stPmsPublish.Header.TimeStamp     := sTimeStamp;

g_stPcsPublish.Header.HeaderVersion := GVL_MQTT.HEADER_VERSION;
g_stPcsPublish.Header.DeviceVersion := GVL_MQTT.DEVICE_VERSION;
g_stPcsPublish.Header.SiteId        := i_stSet.nSiteId;
g_stPcsPublish.Header.DeviceCount   := UINT_TO_UDINT(GVL_PARAM.PCS_COUNT);
g_stPcsPublish.Header.TimeStamp     := sTimeStamp;

g_stBatPublish.Header.HeaderVersion := GVL_MQTT.HEADER_VERSION;
g_stBatPublish.Header.DeviceVersion := GVL_MQTT.DEVICE_VERSION;
g_stBatPublish.Header.SiteId        := i_stSet.nSiteId;
g_stBatPublish.Header.DeviceCount   := UINT_TO_UDINT(GVL_PARAM.BMS_COUNT);
g_stBatPublish.Header.TimeStamp     := sTimeStamp;

g_stRackPublish.Header.HeaderVersion :=GVL_MQTT.HEADER_VERSION;
g_stRackPublish.Header.DeviceVersion := GVL_MQTT.DEVICE_VERSION;
g_stRackPublish.Header.SiteId        := i_stSet.nSiteId;
g_stRackPublish.Header.DeviceCount   := UINT_TO_UDINT(GVL_PARAM.RACK_COUNT);
g_stRackPublish.Header.TimeStamp     := sTimeStamp;

g_stPvPublish.Header.HeaderVersion :=GVL_MQTT.HEADER_VERSION;
g_stPvPublish.Header.DeviceVersion := GVL_MQTT.DEVICE_VERSION;
g_stPvPublish.Header.SiteId        := i_stSet.nSiteId;
g_stPvPublish.Header.DeviceCount   := UINT_TO_UDINT(GVL_PARAM.PV_COUNT);
g_stPvPublish.Header.TimeStamp     := sTimeStamp;

g_stEssPublish.Header.HeaderVersion :=GVL_MQTT.HEADER_VERSION;
g_stEssPublish.Header.DeviceVersion := GVL_MQTT.DEVICE_VERSION;
g_stEssPublish.Header.SiteId        := i_stSet.nSiteId;
g_stEssPublish.Header.DeviceCount   := UINT_TO_UDINT(GVL_PARAM.ESS_COUNT);
g_stEssPublish.Header.TimeStamp     := sTimeStamp;

g_stTempPublish.Header.HeaderVersion :=GVL_MQTT.HEADER_VERSION;
g_stTempPublish.Header.DeviceVersion := GVL_MQTT.DEVICE_VERSION;
g_stTempPublish.Header.SiteId        := i_stSet.nSiteId;
g_stTempPublish.Header.DeviceCount   := UINT_TO_UDINT(GVL_PARAM.TEMP_COUNT);
g_stTempPublish.Header.TimeStamp     := sTimeStamp;

g_stAirConditionerPublish.Header.HeaderVersion := GVL_MQTT.HEADER_VERSION;
g_stAirConditionerPublish.Header.DeviceVersion := GVL_MQTT.DEVICE_VERSION;
g_stAirConditionerPublish.Header.SiteId        := i_stSet.nSiteId;
g_stAirConditionerPublish.Header.DeviceCount   := UINT_TO_UDINT(GVL_PARAM.AIR_CONDITIONER_COUNT);
g_stAirConditionerPublish.Header.TimeStamp     := sTimeStamp;

g_stUpsPublish.Header.HeaderVersion:=GVL_MQTT.HEADER_VERSION;
g_stUpsPublish.Header.DeviceVersion:=GVL_MQTT.DEVICE_VERSION;
g_stUpsPublish.Header.SiteId:=i_stSet.nSiteId;
g_stUpsPublish.Header.DeviceCount:=UINT_TO_UDINT(GVL_PARAM.UPS_COUNT);
g_stUpsPublish.Header.TimeStamp:=sTimeStamp;
g_stModulePublish.Header.HeaderVersion:=GVL_MQTT.HEADER_VERSION;
g_stModulePublish.Header.DeviceVersion:=GVL_MQTT.DEVICE_VERSION;
g_stModulePublish.Header.SiteId:=i_stSet.nSiteId;
g_stModulePublish.Header.DeviceCount:=UINT_TO_UDINT(GVL_PARAM.BAT_MODULE_COUNT);
g_stModulePublish.Header.TimeStamp:=sTimeStamp;
g_stImdPublish.Header.HeaderVersion:=GVL_MQTT.HEADER_VERSION;
g_stImdPublish.Header.DeviceVersion:=GVL_MQTT.DEVICE_VERSION;
g_stImdPublish.Header.SiteId:=i_stSet.nSiteId;
g_stImdPublish.Header.DeviceCount:=UINT_TO_UDINT(GVL_PARAM.IMD_COUNT);
g_stImdPublish.Header.TimeStamp:=sTimeStamp;
g_stFirePublish.Header.HeaderVersion:=GVL_MQTT.HEADER_VERSION;
g_stFirePublish.Header.DeviceVersion:=GVL_MQTT.DEVICE_VERSION;
g_stFirePublish.Header.SiteId:=i_stSet.nSiteId;
g_stFirePublish.Header.DeviceCount:=UINT_TO_UDINT(GVL_PARAM.FIRE_COUNT);
g_stFirePublish.Header.TimeStamp:=sTimeStamp;
g_stUpsConfigEcho.Header.HeaderVersion:=GVL_MQTT.HEADER_VERSION;
g_stUpsConfigEcho.Header.CommandVersion:=GVL_MQTT.COMMAND_VERSION;
g_stUpsConfigEcho.Header.DeviceCount:=UINT_TO_UDINT(GVL_PARAM.UPS_COUNT);
g_stUpsConfigEcho.Header.SiteID:=i_stSet.nSiteId;
g_stUpsConfigEcho.Header.Location:=g_stUpsConfigWireIn.Header.Location;
g_stUpsConfigEcho.Header.UserName:=g_stUpsConfigWireIn.Header.UserName;
g_stUpsConfigEcho.Header.TimeStamp:=sTimeStamp;
MEMCPY(destAddr:=ADR(g_stUpsConfigEcho.Records),srcAddr:=ADR(g_astUpsConfig),n:=SIZEOF(g_astUpsConfig));

(* --- config echo (PCS) --- *)
g_stPcsConfigEcho.Header.HeaderVersion  := GVL_MQTT.HEADER_VERSION;
g_stPcsConfigEcho.Header.CommandVersion := GVL_MQTT.COMMAND_VERSION;
g_stPcsConfigEcho.Header.DeviceCount    := UINT_TO_UDINT(GVL_PARAM.PCS_COUNT);
g_stPcsConfigEcho.Header.Location       := g_stPcsConfigWireIn.Header.Location;	// 받은 값 그대로
g_stPcsConfigEcho.Header.SiteID         := i_stSet.nSiteId;
g_stPcsConfigEcho.Header.UserName       := g_stPcsConfigWireIn.Header.UserName;	// 받은 값 그대로
g_stPcsConfigEcho.Header.TimeStamp      := sTimeStamp;
// [9-21 수정 2026-11-04: 받은 값 대신 실제 반영된 설정을 echo (MAIN FB_EmsConfigApply → GVL_IF → PRG_Mqtt). 아직 없으면 받은 값. 원래 이 줄만:
//   MEMCPY(destAddr := ADR(g_stPcsConfigEcho.Records), srcAddr := ADR(g_astPcsConfig), n := SIZEOF(g_astPcsConfig));]
IF g_bConfigApplied THEN
	MEMCPY(destAddr := ADR(g_stPcsConfigEcho.Records), srcAddr := ADR(g_astPcsConfigApplied), n := SIZEOF(g_astPcsConfigApplied));
ELSE
	MEMCPY(destAddr := ADR(g_stPcsConfigEcho.Records), srcAddr := ADR(g_astPcsConfig), n := SIZEOF(g_astPcsConfig));
END_IF

(* --- config echo (BAT) --- *)
g_stBatConfigEcho.Header.HeaderVersion  := GVL_MQTT.HEADER_VERSION;
g_stBatConfigEcho.Header.CommandVersion := GVL_MQTT.COMMAND_VERSION;
g_stBatConfigEcho.Header.DeviceCount    := UINT_TO_UDINT(GVL_PARAM.BMS_COUNT);
g_stBatConfigEcho.Header.Location       := g_stBatConfigWireIn.Header.Location;
g_stBatConfigEcho.Header.SiteID         := i_stSet.nSiteId;
g_stBatConfigEcho.Header.UserName       := g_stBatConfigWireIn.Header.UserName;
g_stBatConfigEcho.Header.TimeStamp      := sTimeStamp;
// [9-21 수정 2026-11-04: 받은 값 대신 실제 반영된 설정을 echo (MAIN FB_EmsConfigApply → GVL_IF → PRG_Mqtt). 아직 없으면 받은 값. 원래 이 줄만:
//   MEMCPY(destAddr := ADR(g_stBatConfigEcho.Records), srcAddr := ADR(g_astBatConfig), n := SIZEOF(g_astBatConfig));]
IF g_bConfigApplied THEN
	MEMCPY(destAddr := ADR(g_stBatConfigEcho.Records), srcAddr := ADR(g_astBatConfigApplied), n := SIZEOF(g_astBatConfigApplied));
ELSE
	MEMCPY(destAddr := ADR(g_stBatConfigEcho.Records), srcAddr := ADR(g_astBatConfig), n := SIZEOF(g_astBatConfig));
END_IF

(* --- config echo (Protection) --- [결함 12 수정 2026-11-04: 추가] *)
g_stProtectionConfigEcho.Header.HeaderVersion  := GVL_MQTT.HEADER_VERSION;
g_stProtectionConfigEcho.Header.CommandVersion := GVL_MQTT.COMMAND_VERSION;
g_stProtectionConfigEcho.Header.DeviceCount    := 1;
g_stProtectionConfigEcho.Header.Location       := g_stProtectionConfigWireIn.Header.Location;
g_stProtectionConfigEcho.Header.SiteID         := i_stSet.nSiteId;
g_stProtectionConfigEcho.Header.UserName       := g_stProtectionConfigWireIn.Header.UserName;
g_stProtectionConfigEcho.Header.TimeStamp      := sTimeStamp;
g_stProtectionConfigEcho.Record                := g_stProtectionConfig;
END_ACTION

ACTION A_PublishLogger:
(* 로거: 쓰는 브로커마다 다음 이벤트 1건씩 (발생할 때만, QoS 1). 보냈으면 다음 번호로.
   접속이 끊긴 브로커는 큐에 남은 것을 접속한 뒤 이어서 보냄 (LOGGER_QUEUE칸보다 밀리면 fbLogger.q_nLost)
   이중화: Active만 보냄 (i_bPublish, 장치 토픽과 같음). 대기 PLC의 로그는 쌓지 않고 버림:
   Active가 된 뒤 옛 로그를 한꺼번에 보내거나, 두 PLC가 같은 로그를 이중으로 보내지 않게 *)
IF NOT i_bPublish THEN
	anLoggerNext[1] := fbLogger.q_nReceived + 1;
	anLoggerNext[2] := fbLogger.q_nReceived + 1;
	anLoggerNext[3] := fbLogger.q_nReceived + 1;
	RETURN;
END_IF
IF i_stSet.stCloud.bUse THEN
	IF fbLogger.M_GetPacket(i_nSiteId := i_stSet.nSiteId, iq_nNext := anLoggerNext[1], iq_stPacket := stLoggerPacket) THEN
		IF fbCloudPub.M_PublishLogger(i_pPayload := ADR(stLoggerPacket), i_nSize := SIZEOF(stLoggerPacket)) THEN
			anLoggerNext[1] := anLoggerNext[1] + 1;
		END_IF
	END_IF
END_IF
IF i_stSet.stLocal.bUse THEN
	IF fbLogger.M_GetPacket(i_nSiteId := i_stSet.nSiteId, iq_nNext := anLoggerNext[2], iq_stPacket := stLoggerPacket) THEN
		IF fbLocalPub.M_PublishLogger(i_pPayload := ADR(stLoggerPacket), i_nSize := SIZEOF(stLoggerPacket)) THEN
			anLoggerNext[2] := anLoggerNext[2] + 1;
		END_IF
	END_IF
END_IF
IF i_stSet.stAzure.bUse THEN
	IF fbLogger.M_GetPacket(i_nSiteId := i_stSet.nSiteId, iq_nNext := anLoggerNext[3], iq_stPacket := stLoggerPacket) THEN
		IF fbAzurePub.M_PublishLogger(i_pPayload := ADR(stLoggerPacket), i_nSize := SIZEOF(stLoggerPacket)) THEN
			anLoggerNext[3] := anLoggerNext[3] + 1;
		END_IF
	END_IF
END_IF
END_ACTION

ACTION A_MergeRxCount:
(* 브로커 3개 중 어디서든 새로 받은 토픽의 TimeStamp·횟수를 GVL_MQTT에 반영 *)
FOR i := 1 TO GVL_MQTT.COMMAND_TOPIC_COUNT DO
	IF fbCloudSub.q_anCmdRxCount[i] <> anPrevCmdCount[1, i] THEN
		anPrevCmdCount[1, i]	:= fbCloudSub.q_anCmdRxCount[i];
		g_asCmdRxTime[i]		:= fbCloudSub.q_asCmdRxTime[i];
		g_anCmdRxCount[i]		:= g_anCmdRxCount[i] + 1;
	END_IF
	IF fbLocalSub.q_anCmdRxCount[i] <> anPrevCmdCount[2, i] THEN
		anPrevCmdCount[2, i]	:= fbLocalSub.q_anCmdRxCount[i];
		g_asCmdRxTime[i]		:= fbLocalSub.q_asCmdRxTime[i];
		g_anCmdRxCount[i]		:= g_anCmdRxCount[i] + 1;
	END_IF
	IF fbAzureSub.q_anCmdRxCount[i] <> anPrevCmdCount[3, i] THEN
		anPrevCmdCount[3, i]	:= fbAzureSub.q_anCmdRxCount[i];
		g_asCmdRxTime[i]		:= fbAzureSub.q_asCmdRxTime[i];
		g_anCmdRxCount[i]		:= g_anCmdRxCount[i] + 1;
	END_IF
END_FOR
FOR i := 1 TO GVL_MQTT.CONFIG_TOPIC_COUNT DO
	IF fbCloudSub.q_anCfgRxCount[i] <> anPrevCfgCount[1, i] THEN
		anPrevCfgCount[1, i]	:= fbCloudSub.q_anCfgRxCount[i];
		g_asCfgRxTime[i]		:= fbCloudSub.q_asCfgRxTime[i];
		g_anCfgRxRecords[i]		:= fbCloudSub.q_anCfgRxRecords[i];	// [21번 수정 2026-11-09]
		g_anCfgRxCount[i]		:= g_anCfgRxCount[i] + 1;
	END_IF
	IF fbLocalSub.q_anCfgRxCount[i] <> anPrevCfgCount[2, i] THEN
		anPrevCfgCount[2, i]	:= fbLocalSub.q_anCfgRxCount[i];
		g_asCfgRxTime[i]		:= fbLocalSub.q_asCfgRxTime[i];
		g_anCfgRxRecords[i]		:= fbLocalSub.q_anCfgRxRecords[i];	// [21번 수정 2026-11-09]
		g_anCfgRxCount[i]		:= g_anCfgRxCount[i] + 1;
	END_IF
	IF fbAzureSub.q_anCfgRxCount[i] <> anPrevCfgCount[3, i] THEN
		anPrevCfgCount[3, i]	:= fbAzureSub.q_anCfgRxCount[i];
		g_asCfgRxTime[i]		:= fbAzureSub.q_asCfgRxTime[i];
		g_anCfgRxRecords[i]		:= fbAzureSub.q_anCfgRxRecords[i];	// [21번 수정 2026-11-09]
		g_anCfgRxCount[i]		:= g_anCfgRxCount[i] + 1;
	END_IF
END_FOR
END_ACTION

END_FUNCTION_BLOCK

// ---- 20_Module/Mqtt/FB_MqttSubscribe.TcPOU
FUNCTION_BLOCK FB_MqttSubscribe		// MQTT 구독 (브로커 1개): command·config 토픽을 받아 토픽 표대로 수신 배열에 넣고, 토픽별 새 수신을 셈
VAR_INPUT
	i_nSiteId		: UDINT;
	i_sHost			: STRING(15);
	i_nPort			: UINT;
	i_sUserName		: STRING;
	i_sUserPassword	: STRING;	// 접속 값은 첫 호출 때 한 번 읽음
	i_sInstance		: STRING(4) := '';	// ClientId 뒤에 붙임 (이중화: PLC마다 다르게 '-P', '-S'. 같으면 브로커가 서로 끊음)
	i_astCommandTable	: ARRAY[1..GVL_MQTT.COMMAND_TOPIC_COUNT] OF ST_MqttSubEntry;	// FB_MqttMain.A_InitSubscribeTable
	i_astConfigTable	: ARRAY[1..GVL_MQTT.CONFIG_TOPIC_COUNT] OF ST_MqttSubEntry;
END_VAR
VAR_OUTPUT
	q_asCmdRxTime		: ARRAY[1..GVL_MQTT.COMMAND_TOPIC_COUNT] OF STRING(23);	// 토픽별 마지막 헤더 TimeStamp
	q_asCfgRxTime		: ARRAY[1..GVL_MQTT.CONFIG_TOPIC_COUNT] OF STRING(23);
	q_anCmdRxCount		: ARRAY[1..GVL_MQTT.COMMAND_TOPIC_COUNT] OF UDINT;	// 새 수신 횟수 (헤더 TimeStamp가 바뀐 메시지)
	q_anCfgRxCount		: ARRAY[1..GVL_MQTT.CONFIG_TOPIC_COUNT] OF UDINT;
	q_anCfgRxRecords	: ARRAY[1..GVL_MQTT.CONFIG_TOPIC_COUNT] OF UDINT;	// 토픽별 마지막 새 메시지에서 실제로 받은 레코드 수 [21번 수정 2026-11-09: 추가]
	q_bConnected		: BOOL;		// 브로커에 접속됨 (FB_IotMqttClient.bConnected) [9번 수정 2026-11-09: 추가]
END_VAR
VAR
	_sSiteId			: STRING;
	_sClientId			: STRING;
	_sHost				: STRING(15);
	_nPort				: UINT;
	_sUserName			: STRING;
	_sUserPassword		: STRING;
	_asCommandTopic		: ARRAY[1..GVL_MQTT.COMMAND_TOPIC_COUNT] OF STRING(80);
	_asConfigTopic		: ARRAY[1..GVL_MQTT.CONFIG_TOPIC_COUNT] OF STRING(80);
	_fbClient			: FB_IotMqttClient;
	_fbQueue			: FB_IotMqttMessageQueue;
	_fbMessage			: FB_IotMqttMessage;
	_i					: UINT;
	_bSetParameter		: BOOL := TRUE;
	_bConnect			: BOOL := TRUE;
	_bSubscribed		: BOOL;		// 모든 토픽 구독 완료. 연결이 끊기면 지워서 다시 연결되면 다시 구독
	_pHeader			: POINTER TO ST_MqttCommandHeader;
	_nCopied			: UDINT;
	_nReceived			: UDINT;	// 받은 레코드 수 (F_MqttDistribute.q_nReceived)
END_VAR

IF _bSetParameter THEN
	_bSetParameter := FALSE;
	_sSiteId		:= UDINT_TO_STRING(i_nSiteId);
	_sHost			:= i_sHost;
	_nPort			:= i_nPort;
	_sClientId		:= CONCAT(CONCAT('dgsems/sub/', _sSiteId), i_sInstance);
	_sUserName		:= i_sUserName;
	_sUserPassword	:= i_sUserPassword;
	(* dgsems/{solution}/{site_id}/{command|config}/{device_name} *)
	FOR _i := 1 TO GVL_MQTT.COMMAND_TOPIC_COUNT DO
		_asCommandTopic[_i] := CONCAT(CONCAT(CONCAT('dgsems/', GVL_MQTT.SOLUTION_NAME), CONCAT('/', _sSiteId)),
									CONCAT(CONCAT('/', i_astCommandTable[_i].sCategory), CONCAT('/', i_astCommandTable[_i].sTopic)));
	END_FOR
	FOR _i := 1 TO GVL_MQTT.CONFIG_TOPIC_COUNT DO
		_asConfigTopic[_i] := CONCAT(CONCAT(CONCAT('dgsems/', GVL_MQTT.SOLUTION_NAME), CONCAT('/', _sSiteId)),
									CONCAT(CONCAT('/', i_astConfigTable[_i].sCategory), CONCAT('/', i_astConfigTable[_i].sTopic)));
	END_FOR
	_fbClient.sClientId		:= _sClientId;
	_fbClient.sUserName		:= _sUserName;
	_fbClient.sUserPassword	:= _sUserPassword;
	_fbClient.sHostName		:= _sHost;
	_fbClient.nHostPort		:= _nPort;
	_fbClient.sTopicPrefix	:= '';
	_fbClient.ipMessageQueue := _fbQueue;
END_IF

_fbClient.Execute(_bConnect);
q_bConnected := _fbClient.bConnected;	// [9번 수정 2026-11-09: 추가]

(* 구독: 모든 토픽이 성공할 때까지 매 스캔 시도. 연결이 끊기면 다시 구독 *)
IF NOT _fbClient.bConnected THEN
	_bSubscribed := FALSE;
ELSIF NOT _bSubscribed THEN
	_bSubscribed := TRUE;
	FOR _i := 1 TO GVL_MQTT.COMMAND_TOPIC_COUNT DO
		_bSubscribed := _fbClient.Subscribe(sTopic := _asCommandTopic[_i], eQos := TcIotMqttQos.AtMostOnceDelivery) AND _bSubscribed;
	END_FOR
	FOR _i := 1 TO GVL_MQTT.CONFIG_TOPIC_COUNT DO
		_bSubscribed := _fbClient.Subscribe(sTopic := _asConfigTopic[_i], eQos := TcIotMqttQos.AtMostOnceDelivery) AND _bSubscribed;
	END_FOR
END_IF

(* 수신: 한 스캔에 1개 *)
IF _fbQueue.nQueuedMessages > 0 THEN
	IF _fbQueue.Dequeue(fbMessage := _fbMessage) THEN
		FOR _i := 1 TO GVL_MQTT.COMMAND_TOPIC_COUNT DO
			IF _fbMessage.CompareTopic(sTopic := _asCommandTopic[_i]) THEN
				_nCopied := F_MqttDistribute(iq_fbMessage := _fbMessage, iq_stEntry := i_astCommandTable[_i]);
				_pHeader := i_astCommandTable[_i].pRxBuffer;
				IF _nCopied > 0 AND _pHeader <> 0 THEN
					IF _pHeader^.TimeStamp <> q_asCmdRxTime[_i] THEN
						q_asCmdRxTime[_i]	:= _pHeader^.TimeStamp;
						q_anCmdRxCount[_i]	:= q_anCmdRxCount[_i] + 1;
					END_IF
				END_IF
				EXIT;
			END_IF
		END_FOR
		FOR _i := 1 TO GVL_MQTT.CONFIG_TOPIC_COUNT DO
			IF _fbMessage.CompareTopic(sTopic := _asConfigTopic[_i]) THEN
				_nCopied := F_MqttDistribute(iq_fbMessage := _fbMessage, iq_stEntry := i_astConfigTable[_i], q_nReceived => _nReceived);
				_pHeader := i_astConfigTable[_i].pRxBuffer;
				IF _nCopied > 0 AND _pHeader <> 0 THEN
					IF _pHeader^.TimeStamp <> q_asCfgRxTime[_i] THEN
						q_asCfgRxTime[_i]	:= _pHeader^.TimeStamp;
						q_anCfgRxRecords[_i]	:= _nReceived;
						q_anCfgRxCount[_i]	:= q_anCfgRxCount[_i] + 1;
					END_IF
				END_IF
				EXIT;
			END_IF
		END_FOR
	END_IF
END_IF

END_FUNCTION_BLOCK

// ---- 20_Module/Mqtt/F_MqttDistribute.TcPOU
FUNCTION F_MqttDistribute : UDINT		// 받은 MQTT 메시지(헤더 + 레코드 n개)를 토픽 표대로 수신 배열 칸에 복사. 반환 = 복사한 레코드 수
VAR_IN_OUT
	iq_fbMessage	: FB_IotMqttMessage;
	iq_stEntry		: ST_MqttSubEntry;		// 토픽 표 한 칸 (수신 버퍼·목적지·레코드 크기)
END_VAR
VAR_OUTPUT
	q_nReceived		: UDINT;				// 이 메시지에서 실제로 받은 레코드 수 (UPS: 헤더 DeviceCount만큼 다 받았을 때만 그 수, 아니면 0). [21번 수정 2026-11-09: 추가]
END_VAR
VAR CONSTANT
	DEVICE_ID_BASE	: UDINT := 1;			// 받은 레코드의 DeviceIndex(DeviceId) 시작 번호. 모든 command·config 토픽 1부터 (발행 번호와 같음) [1부터 2026-11-10]. 원래 0
END_VAR
VAR
	pHeader			: POINTER TO ST_MqttCommandHeader;
	pRecord			: POINTER TO BYTE;
	pIndex			: POINTER TO UDINT;
	pDest			: POINTER TO BYTE;
	nPayloadBytes	: UDINT;			// 받은 메시지 길이 (byte)
	nRequiredBytes	: UDINT;			// 헤더 DeviceCount에 필요한 길이 (byte)
	nRecords		: UDINT;
	nDev			: UDINT;
	k				: UDINT;
END_VAR

q_nReceived := 0;
// [UPS] 수신 버퍼·목적지·레코드 크기가 없으면, 또는 메시지가 헤더보다 짧거나 수신 버퍼보다 크면 버퍼를 건드리지 않고 버림 (STD 결함 11 수정과 같은 목적, UPS가 더 엄격)
IF iq_stEntry.pRxBuffer=0 OR iq_stEntry.pDestArray=0 OR iq_stEntry.nElementSize=0 THEN RETURN; END_IF
nPayloadBytes:=iq_fbMessage.nPayloadSize;
IF nPayloadBytes<SIZEOF(ST_MqttCommandHeader) OR nPayloadBytes>iq_stEntry.nRxBufferSize THEN RETURN; END_IF
// [STD 9-21 수정 2026-11-04: 받기 전에 수신 버퍼를 0으로 (지난 메시지 레코드가 남지 않게)]
MEMSET(destAddr := iq_stEntry.pRxBuffer, fillByte := 0, n := iq_stEntry.nRxBufferSize);
IF NOT iq_fbMessage.GetPayload(pPayload := iq_stEntry.pRxBuffer, nPayloadSize := iq_stEntry.nRxBufferSize, bSetNullTermination := FALSE) THEN RETURN; END_IF

